// ---- SelfTests/TestCases/TestSuite_CommandAdapter/Test_CommandAdapterInitialization.TcPOU
{region 'Documentation'}
(*!
<summary>Verifies command-only initialization before cyclic use and after a retained sample.</summary>
<description>
PrimeHistory selects the reinitialization case: one public adapter call establishes TRUE history
before Initialize. The other instance calls Initialize before its first-ever cyclic use.
Both variants seed every command and distinctive Name/Status values. Initialize must clear
commands without touching the projection or invoking owner requests. Two fresh samples then
prove the old history was discarded and normal forwarding still works. No Event Buffer is
bound to this request-only double or to the production adapter; buffer work is outside its API.
Repeat runs reinitialize the same instance before the next script, rather than claiming fresh
instance memory. Assertions use the outer selftest publisher; the subject has no publisher.
</description>
*)
{endregion}
FUNCTION_BLOCK Test_CommandAdapterInitialization EXTENDS TestCaseBase
VAR_INPUT
    PrimeHistory : BOOL := FALSE; //! TRUE primes one TRUE command sample before reinitialization; FALSE exercises first-ever initialization.
END_VAR
VAR
    FSubject : RunControlCommandAdapter;
    FOwner : RunControlRequestRecorder;
    FControl : ST_RunControl;
    FExpectedStatus : ST_RunControlStatus;
    FStep : UINT;
    FChecked : BOOL;
    FCommandsCleared : AssertTrue;
    FCommandsClearedMatches : BOOL;
    FProjectionPreserved : AssertTrue;
    FProjectionPreservedMatches : BOOL;
    FNoRequests : AssertTrue;
    FNoRequestsMatches : BOOL;
    FHistoryCleared : AssertTrue;
    FHistoryClearedMatches : BOOL;
    FFreshRequest : AssertTrue;
    FFreshRequestMatches : BOOL;
END_VAR
VAR CONSTANT
    InitializeSubject : UINT := 0;
    FirstSample : UINT := 1;
    SecondSample : UINT := 2;
    CheckResults : UINT := 3;
END_VAR

SUPER^();

{region 'Documentation'}
(*!
<summary>Collects the five independent initialization checks.</summary>
*)
{endregion}
METHOD PROTECTED AggregateResults
VAR_INPUT
    Aggregator : I_ResultAggregator; //! Borrowed result sink owned by the outer Test Case; add this test's checking Assertions without resetting or retaining the sink.
END_VAR
Aggregator.AddProvider(Provider := FCommandsCleared);
Aggregator.AddProvider(Provider := FProjectionPreserved);
Aggregator.AddProvider(Provider := FNoRequests);
Aggregator.AddProvider(Provider := FHistoryCleared);
Aggregator.AddProvider(Provider := FFreshRequest);
END_METHOD

{region 'Documentation'}
(*!
<summary>Configures one scripted initialization test and its checking Assertions.</summary>
*)
{endregion}
METHOD PROTECTED Configure
FPreparationStateCount := 0;
FTestStateCount := 1;
FCommandsCleared.Initialize(Parent := THIS^,
    AssertionName := 'CommandsCleared');
FProjectionPreserved.Initialize(Parent := THIS^,
    AssertionName := 'ProjectionPreserved');
FNoRequests.Initialize(Parent := THIS^,
    AssertionName := 'NoRequests');
FHistoryCleared.Initialize(Parent := THIS^,
    AssertionName := 'HistoryCleared');
FFreshRequest.Initialize(Parent := THIS^,
    AssertionName := 'FreshRequest');
END_METHOD

{region 'Documentation'}
(*!
<summary>No asynchronous resource needs abort processing.</summary>
*)
{endregion}
METHOD PROTECTED ProcessAbort
VAR_INPUT
    Enable : BOOL; //! Phase permission supplied by the owning Test Case; FALSE does not authorize progression, while observation may continue.
END_VAR
IF Enable THEN
    CompleteAbort();
END_IF;
END_METHOD

{region 'Documentation'}
(*!
<summary>Evaluates stored observations after the bounded three-step script.</summary>
*)
{endregion}
METHOD PROTECTED ProcessAssertions
VAR_INPUT
    Enable : BOOL; //! Phase permission supplied by the owning Test Case; FALSE does not authorize progression, while observation may continue.
END_VAR
VAR
    Evaluate : BOOL;
END_VAR
Evaluate := Enable AND (FStep = CheckResults);
FCommandsCleared(Enable := Evaluate,
    State := State,
    IN := FCommandsClearedMatches);
FProjectionPreserved(Enable := Evaluate,
    State := State,
    IN := FProjectionPreservedMatches);
FNoRequests(Enable := Evaluate,
    State := State,
    IN := FNoRequestsMatches);
FHistoryCleared(Enable := Evaluate,
    State := State,
    IN := FHistoryClearedMatches);
FFreshRequest(Enable := Evaluate,
    State := State,
    IN := FFreshRequestMatches);
IF Evaluate THEN
    FChecked := TRUE;
END_IF;
END_METHOD

{region 'Documentation'}
(*!
<summary>No Preparation phase is needed.</summary>
*)
{endregion}
METHOD PROTECTED ProcessPreparations
VAR_INPUT
    // SA0033: Required override; this test has no Preparation work.
    {attribute 'analysis' := '-33'}
    Enable : BOOL; //! Phase permission supplied by the owning Test Case; FALSE does not authorize progression, while observation may continue.
END_VAR
END_METHOD

{region 'Documentation'}
(*!
<summary>Resets the test script; subject initialization remains the operation under test.</summary>
*)
{endregion}
METHOD PROTECTED ProcessReset
FStep := InitializeSubject;
FChecked := FALSE;
FOwner.Clear();
FCommandsCleared.Reset();
FCommandsClearedMatches := FALSE;
FProjectionPreserved.Reset();
FProjectionPreservedMatches := FALSE;
FNoRequests.Reset();
FNoRequestsMatches := FALSE;
FHistoryCleared.Reset();
FHistoryClearedMatches := FALSE;
FFreshRequest.Reset();
FFreshRequestMatches := FALSE;
CompleteReset();
END_METHOD

{region 'Documentation'}
(*!
<summary>Initializes before cyclic use, then checks history through two fresh samples.</summary>
*)
{endregion}
METHOD PROTECTED ProcessTests
VAR_INPUT
    Enable : BOOL; //! Phase permission supplied by the owning Test Case; FALSE does not authorize progression, while observation may continue.
END_VAR
IF NOT Enable THEN
    RETURN;
END_IF;
IF FChecked THEN
    CompleteTests();
    RETURN;
END_IF;
CASE FStep OF
    InitializeSubject:
        SeedControl();
        FOwner.Clear();
        IF PrimeHistory THEN
            // Establish stale TRUE samples through the public call, never by editing private history.
            FSubject(RunControl := FOwner,
                Commands := FControl.Cmd);
            FNoRequestsMatches := (FOwner.StartCount = 0) AND (FOwner.AbortCount = 0) AND (FOwner.ResetCount = 0);
        ELSE
            FNoRequestsMatches := TRUE;
        END_IF;
        FSubject.Initialize(ControlData := FControl);
        FCommandsClearedMatches := NOT FControl.Cmd.Start AND NOT FControl.Cmd.Abort AND NOT FControl.Cmd.Reset
            AND NOT FControl.BufferCmd.Reset AND (FControl.BufferCmd.DeleteSequenceId = 0);
        FProjectionPreservedMatches := (FControl.Name = 'PreservedRoot')
            AND (FControl.Status.Execution.State = FExpectedStatus.Execution.State)
            AND (FControl.Status.Execution.ExecutionStatus = FExpectedStatus.Execution.ExecutionStatus)
            AND (FControl.Status.Execution.Result = FExpectedStatus.Execution.Result)
            AND (FControl.Status.Execution.Uninitialized = FExpectedStatus.Execution.Uninitialized)
            AND (FControl.Status.Execution.ConfigError = FExpectedStatus.Execution.ConfigError)
            AND (FControl.Status.Execution.Ready = FExpectedStatus.Execution.Ready)
            AND (FControl.Status.Execution.Running = FExpectedStatus.Execution.Running)
            AND (FControl.Status.Execution.Completed = FExpectedStatus.Execution.Completed)
            AND (FControl.Status.Execution.Aborted = FExpectedStatus.Execution.Aborted)
            AND (FControl.Status.Execution.Inactive = FExpectedStatus.Execution.Inactive)
            AND (FControl.Status.Execution.Error = FExpectedStatus.Execution.Error)
            AND (FControl.Status.SuiteCountTotal = FExpectedStatus.SuiteCountTotal)
            AND (FControl.Status.SuiteCountInactive = FExpectedStatus.SuiteCountInactive)
            AND (FControl.Status.SuiteCountIdle = FExpectedStatus.SuiteCountIdle)
            AND (FControl.Status.SuiteCountRunning = FExpectedStatus.SuiteCountRunning)
            AND (FControl.Status.SuiteCountCompleted = FExpectedStatus.SuiteCountCompleted)
            AND (FControl.Status.SuiteCountPassed = FExpectedStatus.SuiteCountPassed)
            AND (FControl.Status.SuiteCountFailed = FExpectedStatus.SuiteCountFailed)
            AND (FControl.Status.SuiteCountError = FExpectedStatus.SuiteCountError)
            AND (FControl.Status.Runtime = FExpectedStatus.Runtime);
        FNoRequestsMatches := FNoRequestsMatches AND (FOwner.StartCount = 0) AND (FOwner.AbortCount = 0) AND (FOwner.ResetCount = 0);
        FStep := FirstSample;
    FirstSample:
        FControl.Cmd.Start := TRUE;
        FControl.Cmd.Abort := TRUE;
        FControl.Cmd.Reset := TRUE;
        FSubject(RunControl := FOwner,
            Commands := FControl.Cmd);
        FHistoryClearedMatches := (FOwner.StartCount = 0) AND (FOwner.AbortCount = 0) AND (FOwner.ResetCount = 0)
            AND FControl.Cmd.Start AND FControl.Cmd.Abort AND FControl.Cmd.Reset;
        FStep := SecondSample;
    SecondSample:
        FSubject(RunControl := FOwner,
            Commands := FControl.Cmd);
        FFreshRequestMatches := (FOwner.StartCount = 1) AND (FOwner.AbortCount = 1)
            AND (FOwner.ResetCount = 1) AND NOT FControl.Cmd.Start AND NOT FControl.Cmd.Abort AND NOT FControl.Cmd.Reset;
        FStep := CheckResults;
END_CASE;
END_METHOD

{region 'Documentation'}
(*!
<summary>Uses distinctive projection sentinels, deliberately not a valid lifecycle snapshot.</summary>
*)
{endregion}
METHOD PRIVATE SeedControl
FControl.Name := 'PreservedRoot';
FControl.Status.Execution.State := E_State.Completed;
FControl.Status.Execution.ExecutionStatus := E_ExecutionStatus.Completed;
FControl.Status.Execution.Result := E_Result.Failed;
FControl.Status.Execution.Uninitialized := TRUE;
FControl.Status.Execution.ConfigError := TRUE;
FControl.Status.Execution.Ready := TRUE;
FControl.Status.Execution.Running := TRUE;
FControl.Status.Execution.Completed := TRUE;
FControl.Status.Execution.Aborted := TRUE;
FControl.Status.Execution.Inactive := TRUE;
FControl.Status.Execution.Error := TRUE;
FControl.Status.SuiteCountTotal := 1;
FControl.Status.SuiteCountInactive := 2;
FControl.Status.SuiteCountIdle := 3;
FControl.Status.SuiteCountRunning := 4;
FControl.Status.SuiteCountCompleted := 5;
FControl.Status.SuiteCountPassed := 6;
FControl.Status.SuiteCountFailed := 7;
FControl.Status.SuiteCountError := 8;
FControl.Status.Runtime := T#123ms;
FExpectedStatus := FControl.Status;
FControl.Cmd.Start := TRUE;
FControl.Cmd.Abort := TRUE;
FControl.Cmd.Reset := TRUE;
FControl.BufferCmd.Reset := TRUE;
FControl.BufferCmd.DeleteSequenceId := 123;
END_METHOD

END_FUNCTION_BLOCK

// ---- Framework/RunControl/POU/RunControlCommandAdapter.TcPOU
{region 'Documentation'}
(*!
<summary>Qualifies external lifecycle commands and forwards requests before the Run Control FB call.</summary>
<description>
Initialize with the selected ControlData at PLC startup before the first cyclic call.
Requires a valid Run Control interface and its actual command storage, with stable cyclic wiring.

Call once before the matching concrete Run Control in the same task. A lifecycle bit must be TRUE in two consecutive adapter samples before it is forwarded and cleared. Multiple accepted bits are all forwarded; Run Control later applies Reset over Abort over Start. Initialize clears both lifecycle and Buffer commands at startup, while regular calls handle only lifecycle bits. There is no null-interface check or automatic storage-identity validation; the application owns valid, stable wiring.
</description>
*)
{endregion}
FUNCTION_BLOCK RunControlCommandAdapter
VAR_INPUT
    // SA0027: Parameter denotes the supplied owner interface, not the concrete RunControl FB.
    {attribute 'analysis' := '-27'}
    RunControl : I_RunControl; //! Nonzero request recipient matching Commands storage; an uninitialized owner discards forwarded requests.
END_VAR
VAR_IN_OUT
    Commands : ST_Command; //! Actual external lifecycle-command storage; commands are qualified, forwarded and cleared in place.
END_VAR
VAR
    FPreviousCommands : ST_Command;
END_VAR

IF Commands.Reset AND FPreviousCommands.Reset THEN
    RunControl.RequestReset();
    Commands.Reset := FALSE;
END_IF;

IF Commands.Abort AND FPreviousCommands.Abort THEN
    RunControl.RequestAbort();
    Commands.Abort := FALSE;
END_IF;

IF Commands.Start AND FPreviousCommands.Start THEN
    RunControl.RequestStart();
    Commands.Start := FALSE;
END_IF;

FPreviousCommands := Commands;

{region 'Documentation'}
(*!
<summary>Clears external commands and sampling history once at PLC startup, before Event Buffer/hierarchy initialization.</summary>
<description>
Preserves Name and Status; does not use cyclic inputs, invoke requests or execute buffer operations.
</description>
*)
{endregion}
METHOD PUBLIC Initialize
VAR_IN_OUT
    ControlData : ST_RunControl; //! External Run Control storage; Initialize clears Cmd and BufferCmd without changing Name or Status.
END_VAR
ControlData.Cmd.Start := FALSE;
ControlData.Cmd.Abort := FALSE;
ControlData.Cmd.Reset := FALSE;
ControlData.BufferCmd.Reset := FALSE;
ControlData.BufferCmd.DeleteSequenceId := 0;

FPreviousCommands.Start := FALSE;
FPreviousCommands.Abort := FALSE;
FPreviousCommands.Reset := FALSE;
END_METHOD

END_FUNCTION_BLOCK

// ---- SelfTests/TestCases/TestSuite_CommandAdapter/Helper/RunControlRequestRecorder.TcPOU
{region 'Documentation'}
(*!
<summary>Request-only I_RunControl double; counts calls without simulating lifecycle behavior.</summary>
*)
{endregion}
FUNCTION_BLOCK RunControlRequestRecorder IMPLEMENTS I_RunControl
VAR
    FStartCount : UINT;
    FAbortCount : UINT;
    FResetCount : UINT;
    FStatus : ST_RunControlStatus;
END_VAR

{region 'Documentation'}
(*!
<summary>Passive AbortCount observation for the command-adapter tests.</summary>
*)
{endregion}
{attribute 'monitoring' := 'call'}
PROPERTY PUBLIC AbortCount : UINT //! Passive AbortCount observation for the command-adapter tests.
GET // PUBLIC
AbortCount := FAbortCount;
END_GET
END_PROPERTY

{region 'Documentation'}
(*!
<summary>Clears recorded calls without performing lifecycle work.</summary>
*)
{endregion}
METHOD PUBLIC Clear
FStartCount := 0;
FAbortCount := 0;
FResetCount := 0;
END_METHOD

{region 'Documentation'}
(*!
<summary>Passive Name observation for the command-adapter tests.</summary>
*)
{endregion}
{attribute 'monitoring' := 'variable'}
PROPERTY PUBLIC Name : STRING(GVL_Constants.NameLength) //! Passive Name observation for the command-adapter tests.
GET // PUBLIC
Name := 'CommandTarget';
END_GET
END_PROPERTY

{region 'Documentation'}
(*!
<summary>Records a Abort request only; no lifecycle or buffer operations.</summary>
*)
{endregion}
METHOD PUBLIC RequestAbort
FAbortCount := FAbortCount + 1;
END_METHOD

{region 'Documentation'}
(*!
<summary>Records a Reset request only; no lifecycle or buffer operations.</summary>
*)
{endregion}
METHOD PUBLIC RequestReset
FResetCount := FResetCount + 1;
END_METHOD

{region 'Documentation'}
(*!
<summary>Records a Start request only; no lifecycle or buffer operations.</summary>
*)
{endregion}
METHOD PUBLIC RequestStart
FStartCount := FStartCount + 1;
END_METHOD

{region 'Documentation'}
(*!
<summary>Passive ResetCount observation for the command-adapter tests.</summary>
*)
{endregion}
{attribute 'monitoring' := 'call'}
PROPERTY PUBLIC ResetCount : UINT //! Passive ResetCount observation for the command-adapter tests.
GET // PUBLIC
ResetCount := FResetCount;
END_GET
END_PROPERTY

{region 'Documentation'}
(*!
<summary>Passive Result observation for the command-adapter tests.</summary>
*)
{endregion}
{attribute 'monitoring' := 'call'}
PROPERTY PUBLIC Result : E_Result //! Passive Result observation for the command-adapter tests.
GET // PUBLIC
Result := E_Result.NotEvaluated;
END_GET
END_PROPERTY

{region 'Documentation'}
(*!
<summary>Passive StartCount observation for the command-adapter tests.</summary>
*)
{endregion}
{attribute 'monitoring' := 'call'}
PROPERTY PUBLIC StartCount : UINT //! Passive StartCount observation for the command-adapter tests.
GET // PUBLIC
StartCount := FStartCount;
END_GET
END_PROPERTY

{region 'Documentation'}
(*!
<summary>Passive Status observation for the command-adapter tests.</summary>
*)
{endregion}
PROPERTY PUBLIC Status : ST_RunControlStatus //! Passive Status observation for the command-adapter tests.
GET // PUBLIC
Status := FStatus;
END_GET
END_PROPERTY

END_FUNCTION_BLOCK

// ---- SelfTests/TestCases/TestSuite_CommandAdapter/Test_CommandQualification.TcPOU
{region 'Documentation'}
(*!
<summary>Checks two-sample qualification and PLC-owned clearing for one external lifecycle command.</summary>
<description>
Use one instance per Start, Abort and Reset. Every enabled cycle samples the real adapter once.
The script first withdraws two separate one-sample pulses, then leaves TRUE untouched for two
calls. Acceptance must forward exactly one request and clear that field. A following call
without a write must not repeat it. A new TRUE then needs two new samples before request two.
Each sample checks the selected count/bit and both unrelated commands. This is deterministic
call-boundary evidence, not a simulation of asynchronous ADS writes or a command handshake.
ProcessReset initializes the local subject and clears the recorder for repeatable runs.
</description>
*)
{endregion}
FUNCTION_BLOCK Test_CommandQualification EXTENDS TestCaseBase
VAR_INPUT
    Command : E_AdapterCommand := E_AdapterCommand.Start; //! External command field exercised by this instance; held fixed by the containing Suite.
END_VAR
VAR
    FSubject : RunControlCommandAdapter;
    FOwner : RunControlRequestRecorder;
    FControl : ST_RunControl;
    FStep : UINT;
    FSampleChecked : BOOL;
    FRequestCount : AssertTrue;
    FRequestCountMatches : BOOL;
    FCommandValue : AssertTrue;
    FCommandValueMatches : BOOL;
    FOtherCommands : AssertTrue;
    FOtherCommandsMatches : BOOL;
END_VAR
VAR CONSTANT
    Baseline : UINT := 0;
    SinglePulse : UINT := 1;
    Withdrawal : UINT := 2;
    SeparatedPulse : UINT := 3;
    SecondWithdrawal : UINT := 4;
    RetainedFirstSample : UINT := 5;
    RetainedSecondSample : UINT := 6;
    FreshFirstSample : UINT := 8;
    FreshSecondSample : UINT := 9;
    AfterFreshClearing : UINT := 10;
END_VAR

SUPER^();

{region 'Documentation'}
(*!
<summary>Collects request-count, field-value and isolation checks.</summary>
*)
{endregion}
METHOD PROTECTED AggregateResults
VAR_INPUT
    Aggregator : I_ResultAggregator; //! Borrowed result sink owned by the outer Test Case; add this test's checking Assertions without resetting or retaining the sink.
END_VAR
Aggregator.AddProvider(Provider := FRequestCount);
Aggregator.AddProvider(Provider := FCommandValue);
Aggregator.AddProvider(Provider := FOtherCommands);
END_METHOD

{region 'Documentation'}
(*!
<summary>Checks the explicit script oracle against recorded calls and the post-call command fields.</summary>
*)
{endregion}
METHOD PRIVATE CheckSample
VAR
    ExpectedCount : UINT;
    ExpectedCommand : BOOL;
    ActualCount : UINT;
    ActualCommand : BOOL;
END_VAR
IF FStep >= FreshSecondSample THEN
    ExpectedCount := 2;
ELSIF FStep >= RetainedSecondSample THEN
    ExpectedCount := 1;
END_IF;
ExpectedCommand := (FStep = SinglePulse) OR (FStep = SeparatedPulse)
    OR (FStep = RetainedFirstSample) OR (FStep = FreshFirstSample);
CASE Command OF
    E_AdapterCommand.Start:
        ActualCount := FOwner.StartCount;
        ActualCommand := FControl.Cmd.Start;
        FOtherCommandsMatches := (FOwner.AbortCount = 0) AND (FOwner.ResetCount = 0)
            AND NOT FControl.Cmd.Abort AND NOT FControl.Cmd.Reset;
    E_AdapterCommand.Abort:
        ActualCount := FOwner.AbortCount;
        ActualCommand := FControl.Cmd.Abort;
        FOtherCommandsMatches := (FOwner.StartCount = 0) AND (FOwner.ResetCount = 0)
            AND NOT FControl.Cmd.Start AND NOT FControl.Cmd.Reset;
    E_AdapterCommand.Reset:
        ActualCount := FOwner.ResetCount;
        ActualCommand := FControl.Cmd.Reset;
        FOtherCommandsMatches := (FOwner.StartCount = 0) AND (FOwner.AbortCount = 0)
            AND NOT FControl.Cmd.Start AND NOT FControl.Cmd.Abort;
END_CASE;
FRequestCountMatches := ActualCount = ExpectedCount;
FCommandValueMatches := ActualCommand = ExpectedCommand;
END_METHOD

{region 'Documentation'}
(*!
<summary>Initializes the three checking Assertions for the selected command.</summary>
*)
{endregion}
METHOD PROTECTED Configure
FPreparationStateCount := 0;
FTestStateCount := 1;
FRequestCount.Initialize(Parent := THIS^,
    AssertionName := 'RequestCount');
FCommandValue.Initialize(Parent := THIS^,
    AssertionName := 'CommandValue');
FOtherCommands.Initialize(Parent := THIS^,
    AssertionName := 'OtherCommands');
END_METHOD

{region 'Documentation'}
(*!
<summary>No asynchronous resource needs abort handling.</summary>
*)
{endregion}
METHOD PROTECTED ProcessAbort
VAR_INPUT
    Enable : BOOL; //! Phase permission supplied by the owning Test Case; FALSE does not authorize progression, while observation may continue.
END_VAR
IF Enable THEN
    CompleteAbort();
END_IF;
END_METHOD

{region 'Documentation'}
(*!
<summary>Checks every sample before advancing; failures remain latched across the script.</summary>
*)
{endregion}
METHOD PROTECTED ProcessAssertions
VAR_INPUT
    Enable : BOOL; //! Phase permission supplied by the owning Test Case; FALSE does not authorize progression, while observation may continue.
END_VAR
FRequestCount(Enable := Enable,
    State := State,
    IN := FRequestCountMatches);
FCommandValue(Enable := Enable,
    State := State,
    IN := FCommandValueMatches);
FOtherCommands(Enable := Enable,
    State := State,
    IN := FOtherCommandsMatches);
IF Enable THEN
    FSampleChecked := TRUE;
END_IF;
END_METHOD

{region 'Documentation'}
(*!
<summary>No Preparation work is required.</summary>
*)
{endregion}
METHOD PROTECTED ProcessPreparations
VAR_INPUT
    // SA0033: Required override; this test has no Preparation phase.
    {attribute 'analysis' := '-33'}
    Enable : BOOL; //! Phase permission supplied by the owning Test Case; FALSE does not authorize progression, while observation may continue.
END_VAR
END_METHOD

{region 'Documentation'}
(*!
<summary>Clears subject history, recorded requests and the bounded sample script.</summary>
*)
{endregion}
METHOD PROTECTED ProcessReset
FSubject.Initialize(ControlData := FControl);
FOwner.Clear();
FStep := Baseline;
FSampleChecked := FALSE;
FRequestCount.Reset();
FRequestCountMatches := FALSE;
FCommandValue.Reset();
FCommandValueMatches := FALSE;
FOtherCommands.Reset();
FOtherCommandsMatches := FALSE;
CompleteReset();
END_METHOD

{region 'Documentation'}
(*!
<summary>Applies one scheduled write and one real adapter call per active PLC cycle.</summary>
*)
{endregion}
METHOD PROTECTED ProcessTests
VAR_INPUT
    Enable : BOOL; //! Phase permission supplied by the owning Test Case; FALSE does not authorize progression, while observation may continue.
END_VAR
IF NOT Enable THEN
    RETURN;
END_IF;
IF FSampleChecked THEN
    IF FStep = AfterFreshClearing THEN
        CompleteTests();
        RETURN;
    END_IF;
    FStep := FStep + 1;
    FSampleChecked := FALSE;
END_IF;
CASE FStep OF
    SinglePulse, SeparatedPulse, RetainedFirstSample, FreshFirstSample:
        SetCommand(Value := TRUE);
    Withdrawal, SecondWithdrawal:
        SetCommand(Value := FALSE);
ELSE
    // No external write: retain the actual field, including the adapter's clearing.
END_CASE;
FSubject(RunControl := FOwner,
    Commands := FControl.Cmd);
CheckSample();
END_METHOD

{region 'Documentation'}
(*!
<summary>Writes only the chosen external command field.</summary>
*)
{endregion}
METHOD PRIVATE SetCommand
VAR_INPUT
    Value : BOOL; //! Boolean value written only to the selected command field.
END_VAR
CASE Command OF
    E_AdapterCommand.Start:
        FControl.Cmd.Start := Value;
    E_AdapterCommand.Abort:
        FControl.Cmd.Abort := Value;
    E_AdapterCommand.Reset:
        FControl.Cmd.Reset := Value;
END_CASE;
END_METHOD

END_FUNCTION_BLOCK

// ---- SelfTests/TestCases/TestSuite_CommandAdapter/Test_CommandIndependence.TcPOU
{region 'Documentation'}
(*!
<summary>Verifies independent command qualification and selective clearing across staggered writes.</summary>
<description>
The initial Start/Reset pair is sampled before Abort is written after that call. The pair
must be forwarded while Abort remains pending. Further post-call Start, Reset and Abort
writes rotate which field is newly sampled versus accepted. After those requests drain,
all three bits are raised together and must all be forwarded exactly once after two samples.
Fixed count and bit traces are the oracle; no request order or lifecycle priority is asserted.
Buffer commands and selected Name/Status fields are changed before each call and must survive.
CheckSample captures pre-post-write observations so Assertion processing cannot confuse the
test's own later writes with the adapter's output. There is one subject call per active cycle.
These deterministic boundaries do not prove arbitrary ADS interleavings inside an FB call.
</description>
*)
{endregion}
FUNCTION_BLOCK Test_CommandIndependence EXTENDS TestCaseBase
VAR
    FSubject : RunControlCommandAdapter;
    FOwner : RunControlRequestRecorder;
    FControl : ST_RunControl;
    FStep : UINT;
    FSampleChecked : BOOL;
    FForwarding : AssertTrue;
    FForwardingMatches : BOOL;
    FSelectiveClearing : AssertTrue;
    FSelectiveClearingMatches : BOOL;
    FUnrelatedFields : AssertTrue;
    FUnrelatedFieldsMatches : BOOL;
END_VAR
VAR CONSTANT
    PairFirstSample : UINT := 0;
    PairAccepted : UINT := 1;
    AbortAccepted : UINT := 2;
    StartAccepted : UINT := 3;
    ResetAccepted : UINT := 4;
    SecondAbortAccepted : UINT := 5;
    AllFirstSample : UINT := 8;
    LastSample : UINT := 10;
    ExpectedStartCounts : ARRAY[0..LastSample] OF UINT := [0, 1, 1, 2, 2, 2, 3, 3, 3, 4, 4];
    ExpectedAbortCounts : ARRAY[0..LastSample] OF UINT := [0, 0, 1, 1, 1, 2, 2, 2, 2, 3, 3];
    ExpectedResetCounts : ARRAY[0..LastSample] OF UINT := [0, 1, 1, 1, 2, 2, 2, 3, 3, 4, 4];
    ExpectedStartBits : ARRAY[0..LastSample] OF BOOL := [TRUE, FALSE, TRUE, FALSE, FALSE, TRUE, FALSE, FALSE, TRUE, FALSE, FALSE];
    ExpectedAbortBits : ARRAY[0..LastSample] OF BOOL := [FALSE, TRUE, FALSE, FALSE, TRUE, FALSE, FALSE, FALSE, TRUE, FALSE, FALSE];
    ExpectedResetBits : ARRAY[0..LastSample] OF BOOL := [TRUE, FALSE, FALSE, TRUE, FALSE, FALSE, TRUE, FALSE, TRUE, FALSE, FALSE];
END_VAR

SUPER^();

{region 'Documentation'}
(*!
<summary>Collects only the checking Assertions.</summary>
*)
{endregion}
METHOD PROTECTED AggregateResults
VAR_INPUT
    Aggregator : I_ResultAggregator; //! Borrowed result sink owned by the outer Test Case; add this test's checking Assertions without resetting or retaining the sink.
END_VAR
Aggregator.AddProvider(Provider := FForwarding);
Aggregator.AddProvider(Provider := FSelectiveClearing);
Aggregator.AddProvider(Provider := FUnrelatedFields);
END_METHOD

{region 'Documentation'}
(*!
<summary>Uses fixed expected traces, independent of adapter request order.</summary>
*)
{endregion}
METHOD PRIVATE CheckSample
FForwardingMatches := (FOwner.StartCount = ExpectedStartCounts[FStep])
    AND (FOwner.AbortCount = ExpectedAbortCounts[FStep])
    AND (FOwner.ResetCount = ExpectedResetCounts[FStep]);
FSelectiveClearingMatches := (FControl.Cmd.Start = ExpectedStartBits[FStep])
    AND (FControl.Cmd.Abort = ExpectedAbortBits[FStep])
    AND (FControl.Cmd.Reset = ExpectedResetBits[FStep]);
FUnrelatedFieldsMatches := (FControl.Name = 'CommandProjection')
    AND (FControl.Status.Execution.State = E_State.Completed)
    AND (FControl.Status.Execution.Result = E_Result.Failed)
    AND (FControl.Status.SuiteCountTotal = FStep + 1)
    AND (FControl.Status.Runtime = UINT_TO_TIME(FStep + 1))
    AND (FControl.BufferCmd.Reset = ((FStep MOD 2) = 0))
    AND (FControl.BufferCmd.DeleteSequenceId = UINT_TO_UDINT(FStep + 1));
END_METHOD

{region 'Documentation'}
(*!
<summary>Initializes the independent forwarding, clearing and projection checks.</summary>
*)
{endregion}
METHOD PROTECTED Configure
FPreparationStateCount := 0;
FTestStateCount := 1;
FForwarding.Initialize(Parent := THIS^,
    AssertionName := 'Forwarding');
FSelectiveClearing.Initialize(Parent := THIS^,
    AssertionName := 'SelectiveClearing');
FUnrelatedFields.Initialize(Parent := THIS^,
    AssertionName := 'UnrelatedFields');
END_METHOD

{region 'Documentation'}
(*!
<summary>No asynchronous resource is involved.</summary>
*)
{endregion}
METHOD PROTECTED ProcessAbort
VAR_INPUT
    Enable : BOOL; //! Phase permission supplied by the owning Test Case; FALSE does not authorize progression, while observation may continue.
END_VAR
IF Enable THEN
    CompleteAbort();
END_IF;
END_METHOD

{region 'Documentation'}
(*!
<summary>Latches every sample's observations before the script advances.</summary>
*)
{endregion}
METHOD PROTECTED ProcessAssertions
VAR_INPUT
    Enable : BOOL; //! Phase permission supplied by the owning Test Case; FALSE does not authorize progression, while observation may continue.
END_VAR
FForwarding(Enable := Enable,
    State := State,
    IN := FForwardingMatches);
FSelectiveClearing(Enable := Enable,
    State := State,
    IN := FSelectiveClearingMatches);
FUnrelatedFields(Enable := Enable,
    State := State,
    IN := FUnrelatedFieldsMatches);
IF Enable THEN
    FSampleChecked := TRUE;
END_IF;
END_METHOD

{region 'Documentation'}
(*!
<summary>No Preparation phase is required.</summary>
*)
{endregion}
METHOD PROTECTED ProcessPreparations
VAR_INPUT
    // SA0033: Required override; this test has no Preparation phase.
    {attribute 'analysis' := '-33'}
    Enable : BOOL; //! Phase permission supplied by the owning Test Case; FALSE does not authorize progression, while observation may continue.
END_VAR
END_METHOD

{region 'Documentation'}
(*!
<summary>Clears local commands, sampling history, recorded calls and checking state.</summary>
*)
{endregion}
METHOD PROTECTED ProcessReset
FSubject.Initialize(ControlData := FControl);
FOwner.Clear();
FStep := PairFirstSample;
FSampleChecked := FALSE;
FForwarding.Reset();
FForwardingMatches := FALSE;
FSelectiveClearing.Reset();
FSelectiveClearingMatches := FALSE;
FUnrelatedFields.Reset();
FUnrelatedFieldsMatches := FALSE;
CompleteReset();
END_METHOD

{region 'Documentation'}
(*!
<summary>Places writes before or after one adapter call; captures observations before post-call writes.</summary>
*)
{endregion}
METHOD PROTECTED ProcessTests
VAR_INPUT
    Enable : BOOL; //! Phase permission supplied by the owning Test Case; FALSE does not authorize progression, while observation may continue.
END_VAR
IF NOT Enable THEN
    RETURN;
END_IF;
IF FSampleChecked THEN
    IF FStep = LastSample THEN
        CompleteTests();
        RETURN;
    END_IF;
    FStep := FStep + 1;
    FSampleChecked := FALSE;
END_IF;
CASE FStep OF
    PairFirstSample:
        FControl.Cmd.Start := TRUE;
        FControl.Cmd.Reset := TRUE;
    AllFirstSample:
        FControl.Cmd.Start := TRUE;
        FControl.Cmd.Abort := TRUE;
        FControl.Cmd.Reset := TRUE;
END_CASE;
FControl.Name := 'CommandProjection';
FControl.Status.Execution.State := E_State.Completed;
FControl.Status.Execution.Result := E_Result.Failed;
FControl.Status.SuiteCountTotal := FStep + 1;
FControl.Status.Runtime := UINT_TO_TIME(FStep + 1);
FControl.BufferCmd.Reset := (FStep MOD 2) = 0;
FControl.BufferCmd.DeleteSequenceId := UINT_TO_UDINT(FStep + 1);
FSubject(RunControl := FOwner,
    Commands := FControl.Cmd);
CheckSample();
// These writes happen after the observation and become the next call's first sample.
CASE FStep OF
    PairFirstSample, StartAccepted:
        FControl.Cmd.Abort := TRUE;
    PairAccepted, ResetAccepted:
        FControl.Cmd.Start := TRUE;
    AbortAccepted, SecondAbortAccepted:
        FControl.Cmd.Reset := TRUE;
END_CASE;
END_METHOD

END_FUNCTION_BLOCK

// ---- SelfTests/TestSuites/TestSuite_EventDelivery.TcPOU
{region 'Documentation'}
(*!
<summary>Groups isolated event storage, delivery and deletion-watermark tests.</summary>
*)
{endregion}
FUNCTION_BLOCK TestSuite_EventDelivery EXTENDS TestSuiteBase
VAR
    FStorageBinding : Test_EventStorageBinding;
    FContent : Test_EventContent;
    FBufferFull : Test_EventBufferFull;
    FRingOrder : Test_EventRingOrder;
    FDeleteWatermarks : Test_EventDeleteWatermarks;
    FDeleteWrappedFull : Test_EventDeleteWrappedFull;
    FDeleteLostSequence : Test_EventDeleteLostSequence;
    FDeleteCommandBoundary : Test_EventDeleteCommandBoundary;
    FTestCases : ARRAY[1..TestCaseCapacity] OF I_TestCase;
END_VAR
VAR CONSTANT
    TestCaseCapacity : UINT := 8;
END_VAR

SUPER^();

{region 'Documentation'}
(*!
<summary>Initializes and registers the isolated event scenarios for serial execution.</summary>
*)
{endregion}
METHOD PROTECTED Configure
VAR_IN_OUT
    // SA0167: Borrowed owner builder; no temporary instance is created.
    {attribute 'analysis' := '-167'}
    Builder : TestSuiteConfigurationBuilder; //! Borrowed owner configuration builder used only during this Configure call; register this owner's concrete children.
END_VAR
VAR
    TestConfig : ST_TestCaseConfig;
END_VAR
Builder.Initialize(Mode := E_OrchestrationMode.Serial,
    TestCases := FTestCases);
FStorageBinding.Initialize(Parent := THIS^,
    TestName := 'StorageBinding',
    Config := TestConfig);
Builder.Register(TestCase := FStorageBinding);
FContent.Initialize(Parent := THIS^,
    TestName := 'Content',
    Config := TestConfig);
Builder.Register(TestCase := FContent);
FBufferFull.Initialize(Parent := THIS^,
    TestName := 'BufferFull',
    Config := TestConfig);
Builder.Register(TestCase := FBufferFull);
FRingOrder.Initialize(Parent := THIS^,
    TestName := 'RingOrder',
    Config := TestConfig);
Builder.Register(TestCase := FRingOrder);
FDeleteWatermarks.Initialize(Parent := THIS^,
    TestName := 'DeleteWatermarks',
    Config := TestConfig);
Builder.Register(TestCase := FDeleteWatermarks);
FDeleteWrappedFull.Initialize(Parent := THIS^,
    TestName := 'DeleteWrappedFull',
    Config := TestConfig);
Builder.Register(TestCase := FDeleteWrappedFull);
FDeleteLostSequence.Initialize(Parent := THIS^,
    TestName := 'DeleteLostSequence',
    Config := TestConfig);
Builder.Register(TestCase := FDeleteLostSequence);
FDeleteCommandBoundary.Initialize(Parent := THIS^,
    TestName := 'DeleteCommandBoundary',
    Config := TestConfig);
Builder.Register(TestCase := FDeleteCommandBoundary);
END_METHOD

{region 'Documentation'}
(*!
<summary>Returns a registered scenario using its original array index.</summary>
*)
{endregion}
METHOD PUBLIC GetTestCase : I_TestCase //! Typed child interface at the original array index; zero when no entry is available.
VAR_INPUT
    Index : DINT; //! Original occupied child-array index, rather than an ordinal position.
END_VAR
GetTestCase := 0;
IF (ChildCount = 0) OR (Index < ChildArrayLowerBound)
    OR (DINT_TO_LINT(Index) >= DINT_TO_LINT(ChildArrayLowerBound) + UINT_TO_LINT(ChildCount)) THEN
    RETURN;
END_IF;
GetTestCase := FTestCases[Index];
END_METHOD

{region 'Documentation'}
(*!
<summary>Calls each owned scenario once per initialized Suite cycle.</summary>
*)
{endregion}
METHOD PROTECTED ProcessTestCases
FStorageBinding();
FContent();
FBufferFull();
FRingOrder();
FDeleteWatermarks();
FDeleteWrappedFull();
FDeleteLostSequence();
FDeleteCommandBoundary();
END_METHOD

END_FUNCTION_BLOCK

// ---- SelfTests/TestCases/TestSuite_EventDelivery/Test_EventStorageBinding.TcPOU
{region 'Documentation'}
(*!
<summary>Verifies two real Event Buffers publish into their own bound arrays and status structures.</summary>
<description>
The subjects own no global stream: each binds a static local array and separate projections.
Eight and twelve physical entries provide seven and eleven usable FIFO slots. One distinctive
event is published to each subject; observations are captured before the next operation so
cross-writes cannot be hidden by later initialization. The outer test Assertions use the
normal selftest publisher, which is never replaced. Every test run initializes both subjects
again; no production algorithm is copied and no private field is modified.
</description>
*)
{endregion}
FUNCTION_BLOCK Test_EventStorageBinding EXTENDS TestCaseBase
VAR
    FSmallBuffer : EventBuffer;
    FLargeBuffer : EventBuffer;
    FSmallEvents : ARRAY[1..SmallBufferLength] OF ST_Event;
    FLargeEvents : ARRAY[1..LargeBufferLength] OF ST_Event;
    FSmallFifo : ST_FifoStatus;
    FLargeFifo : ST_FifoStatus;
    FSmallStatus : ST_EventBufferStatus;
    FLargeStatus : ST_EventBufferStatus;
    FPerformed : BOOL;
    FChecked : BOOL;
    FBinding : AssertTrue;
    FBindingMatches : BOOL;
    FCapacity : AssertTrue;
    FCapacityMatches : BOOL;
    FInitialProjection : AssertTrue;
    FInitialProjectionMatches : BOOL;
    FSmallPublication : AssertTrue;
    FSmallPublicationMatches : BOOL;
    FLargePublication : AssertTrue;
    FLargePublicationMatches : BOOL;
    FIsolation : AssertTrue;
    FIsolationMatches : BOOL;
END_VAR
VAR CONSTANT
    SmallBufferLength : UINT := 8;
    LargeBufferLength : UINT := 12;
END_VAR

SUPER^();

{region 'Documentation'}
(*!
<summary>Collects the six independent storage-binding observations.</summary>
*)
{endregion}
METHOD PROTECTED AggregateResults
VAR_INPUT
    Aggregator : I_ResultAggregator; //! Borrowed result sink owned by the outer Test Case; add this test's checking Assertions without resetting or retaining the sink.
END_VAR
Aggregator.AddProvider(Provider := FBinding);
Aggregator.AddProvider(Provider := FCapacity);
Aggregator.AddProvider(Provider := FInitialProjection);
Aggregator.AddProvider(Provider := FSmallPublication);
Aggregator.AddProvider(Provider := FLargePublication);
Aggregator.AddProvider(Provider := FIsolation);
END_METHOD

{region 'Documentation'}
(*!
<summary>Requires successful initialization of all checking Assertions.</summary>
*)
{endregion}
METHOD PROTECTED CheckInitialization : BOOL //! TRUE when the inherited initialization check and this concrete fixture check both accept the setup.
CheckInitialization := FALSE;
IF NOT SUPER^.CheckInitialization() THEN
    RETURN;
END_IF;

CheckInitialization := FBinding.IsInitialized
    AND FCapacity.IsInitialized
    AND FInitialProjection.IsInitialized
    AND FSmallPublication.IsInitialized
    AND FLargePublication.IsInitialized
    AND FIsolation.IsInitialized;
END_METHOD

{region 'Documentation'}
(*!
<summary>Configures the single storage-binding scenario and its six Assertions.</summary>
*)
{endregion}
METHOD PROTECTED Configure
FPreparationStateCount := 0;
FTestStateCount := 1;
FBinding.Initialize(Parent := THIS^,
    AssertionName := 'Binding');
FCapacity.Initialize(Parent := THIS^,
    AssertionName := 'Capacity');
FInitialProjection.Initialize(Parent := THIS^,
    AssertionName := 'InitialProjection');
FSmallPublication.Initialize(Parent := THIS^,
    AssertionName := 'SmallPublication');
FLargePublication.Initialize(Parent := THIS^,
    AssertionName := 'LargePublication');
FIsolation.Initialize(Parent := THIS^,
    AssertionName := 'Isolation');
END_METHOD

{region 'Documentation'}
(*!
<summary>Binds differently sized static arrays and verifies initial projection and usable capacity.</summary>
*)
{endregion}
METHOD PRIVATE InitializeBuffers
VAR
    SmallInitialized : BOOL;
    LargeInitialized : BOOL;
    Index : UINT;
END_VAR
SmallInitialized := FSmallBuffer.Initialize(Buffer := FSmallEvents,
    FifoControl := FSmallFifo,
    Status := FSmallStatus);
LargeInitialized := FLargeBuffer.Initialize(Buffer := FLargeEvents,
    FifoControl := FLargeFifo,
    Status := FLargeStatus);
FBindingMatches := SmallInitialized AND LargeInitialized
    AND FSmallBuffer.IsValid AND FLargeBuffer.IsValid;
FCapacityMatches := (FSmallBuffer.Capacity = SmallBufferLength - 1)
    AND (FLargeBuffer.Capacity = LargeBufferLength - 1)
    AND (FSmallFifo.BufferLength = SmallBufferLength)
    AND (FLargeFifo.BufferLength = LargeBufferLength);
FInitialProjectionMatches := FSmallFifo.BufferEmpty AND FLargeFifo.BufferEmpty
    AND NOT FSmallFifo.ConfigError AND NOT FLargeFifo.ConfigError
    AND NOT FSmallFifo.IndexError AND NOT FLargeFifo.IndexError
    AND (FSmallFifo.ElementCount = 0) AND (FLargeFifo.ElementCount = 0)
    AND (FSmallFifo.IndexIn = 1) AND (FSmallFifo.IndexOut = 1)
    AND (FLargeFifo.IndexIn = 1) AND (FLargeFifo.IndexOut = 1)
    AND (FSmallStatus.SequenceId = 0) AND (FLargeStatus.SequenceId = 0)
    AND (FSmallStatus.DeletedSequenceId = 0) AND (FLargeStatus.DeletedSequenceId = 0)
    AND (FSmallStatus.LostEventCount = 0) AND (FLargeStatus.LostEventCount = 0);
FOR Index := 1 TO SmallBufferLength DO
    FInitialProjectionMatches := FInitialProjectionMatches AND (FSmallEvents[Index].SequenceId = 0);
END_FOR;
FOR Index := 1 TO LargeBufferLength DO
    FInitialProjectionMatches := FInitialProjectionMatches AND (FLargeEvents[Index].SequenceId = 0);
END_FOR;
END_METHOD

{region 'Documentation'}
(*!
<summary>Completes abort without asynchronous resource work.</summary>
*)
{endregion}
METHOD PROTECTED ProcessAbort
VAR_INPUT
    Enable : BOOL; //! Phase permission supplied by the owning Test Case; FALSE does not authorize progression, while observation may continue.
END_VAR
IF Enable THEN
    CompleteAbort();
END_IF;
END_METHOD

{region 'Documentation'}
(*!
<summary>Evaluates observations only after the two subjects have been exercised.</summary>
*)
{endregion}
METHOD PROTECTED ProcessAssertions
VAR_INPUT
    Enable : BOOL; //! Phase permission supplied by the owning Test Case; FALSE does not authorize progression, while observation may continue.
END_VAR
VAR
    Evaluate : BOOL;
END_VAR
Evaluate := Enable AND FPerformed;
FBinding(Enable := Evaluate,
    State := State,
    IN := FBindingMatches);
FCapacity(Enable := Evaluate,
    State := State,
    IN := FCapacityMatches);
FInitialProjection(Enable := Evaluate,
    State := State,
    IN := FInitialProjectionMatches);
FSmallPublication(Enable := Evaluate,
    State := State,
    IN := FSmallPublicationMatches);
FLargePublication(Enable := Evaluate,
    State := State,
    IN := FLargePublicationMatches);
FIsolation(Enable := Evaluate,
    State := State,
    IN := FIsolationMatches);
IF Evaluate THEN
    FChecked := TRUE;
END_IF;
END_METHOD

{region 'Documentation'}
(*!
<summary>No Preparation phase is needed.</summary>
*)
{endregion}
METHOD PROTECTED ProcessPreparations
VAR_INPUT
    // SA0033: Required override; this test has no Preparation work.
    {attribute 'analysis' := '-33'}
    Enable : BOOL; //! Phase permission supplied by the owning Test Case; FALSE does not authorize progression, while observation may continue.
END_VAR
END_METHOD

{region 'Documentation'}
(*!
<summary>Clears observations and Assertions; subject initialization remains under test.</summary>
*)
{endregion}
METHOD PROTECTED ProcessReset
FPerformed := FALSE;
FChecked := FALSE;
FBinding.Reset();
FBindingMatches := FALSE;
FCapacity.Reset();
FCapacityMatches := FALSE;
FInitialProjection.Reset();
FInitialProjectionMatches := FALSE;
FSmallPublication.Reset();
FSmallPublicationMatches := FALSE;
FLargePublication.Reset();
FLargePublicationMatches := FALSE;
FIsolation.Reset();
FIsolationMatches := FALSE;
CompleteReset();
END_METHOD

{region 'Documentation'}
(*!
<summary>Initializes and exercises the local bindings once per test run.</summary>
*)
{endregion}
METHOD PROTECTED ProcessTests
VAR_INPUT
    Enable : BOOL; //! Phase permission supplied by the owning Test Case; FALSE does not authorize progression, while observation may continue.
END_VAR
IF NOT Enable THEN
    RETURN;
END_IF;
IF FChecked THEN
    CompleteTests();
    RETURN;
END_IF;

IF NOT FPerformed THEN
    InitializeBuffers();
    PublishToSmallBuffer();
    PublishToLargeBuffer();
    FPerformed := TRUE;
END_IF;
END_METHOD

{region 'Documentation'}
(*!
<summary>Checks the second publication leaves the first buffer and its projections unchanged.</summary>
*)
{endregion}
METHOD PRIVATE PublishToLargeBuffer
VAR
    WriteResult : INT;
    Index : UINT;
END_VAR
WriteResult := FLargeBuffer.PublishEvent(Event := CreateFrameworkEvent(Name := 'LocalLarge',
    State := E_State.Idle,
    Severity := E_EventSeverity.Info,
    Message := 'Large binding'));
FLargePublicationMatches := (WriteResult = 1)
    AND (FLargeEvents[1].SequenceId = 1)
    AND (FLargeEvents[1].Name = 'LocalLarge') AND (FLargeEvents[1].Message = 'Large binding')
    AND (FLargeFifo.IndexIn = 2) AND (FLargeFifo.IndexOut = 1)
    AND (FLargeFifo.ElementCount = 1) AND NOT FLargeFifo.BufferEmpty
    AND (FLargeStatus.SequenceId = 1) AND (FLargeStatus.DeletedSequenceId = 0)
    AND (FLargeStatus.LostEventCount = 0);
FIsolationMatches := FIsolationMatches
    AND (FSmallEvents[1].SequenceId = 1)
    AND (FSmallEvents[1].Name = 'LocalSmall') AND (FSmallEvents[1].Message = 'Small binding')
    AND (FSmallFifo.IndexIn = 2) AND (FSmallFifo.IndexOut = 1)
    AND (FSmallFifo.ElementCount = 1) AND NOT FSmallFifo.BufferEmpty
    AND (FSmallStatus.SequenceId = 1) AND (FSmallStatus.DeletedSequenceId = 0)
    AND (FSmallStatus.LostEventCount = 0);
FOR Index := 2 TO SmallBufferLength DO
    FIsolationMatches := FIsolationMatches AND (FSmallEvents[Index].SequenceId = 0);
END_FOR;
END_METHOD

{region 'Documentation'}
(*!
<summary>Checks immediate local publication and that the other buffer is still empty.</summary>
*)
{endregion}
METHOD PRIVATE PublishToSmallBuffer
VAR
    WriteResult : INT;
    Index : UINT;
END_VAR
WriteResult := FSmallBuffer.PublishEvent(Event := CreateFrameworkEvent(Name := 'LocalSmall',
    State := E_State.Idle,
    Severity := E_EventSeverity.Info,
    Message := 'Small binding'));
FSmallPublicationMatches := (WriteResult = 1)
    AND (FSmallEvents[1].SequenceId = 1)
    AND (FSmallEvents[1].Name = 'LocalSmall') AND (FSmallEvents[1].Message = 'Small binding')
    AND (FSmallFifo.IndexIn = 2) AND (FSmallFifo.IndexOut = 1)
    AND (FSmallFifo.ElementCount = 1) AND NOT FSmallFifo.BufferEmpty
    AND (FSmallStatus.SequenceId = 1) AND (FSmallStatus.DeletedSequenceId = 0)
    AND (FSmallStatus.LostEventCount = 0);
FIsolationMatches := FLargeFifo.BufferEmpty AND (FLargeFifo.ElementCount = 0)
    AND (FLargeFifo.IndexIn = 1) AND (FLargeFifo.IndexOut = 1)
    AND (FLargeStatus.SequenceId = 0) AND (FLargeStatus.DeletedSequenceId = 0)
    AND (FLargeStatus.LostEventCount = 0);
FOR Index := 1 TO LargeBufferLength DO
    FIsolationMatches := FIsolationMatches AND (FLargeEvents[Index].SequenceId = 0);
END_FOR;
END_METHOD

END_FUNCTION_BLOCK

// ---- SelfTests/TestCases/TestSuite_EventDelivery/Test_EventContent.TcPOU
{region 'Documentation'}
(*!
<summary>Verifies representative event payloads and producer-assigned identity through real publication.</summary>
<description>
Publishes a state transition, a failed Assertion and a Test Case aggregation. Expectations
state the required fields explicitly instead of constructing the expected event with the same FC.
Sequence and timestamp sentinels verify that the publisher assigns identity to its value copy.
Timestamp checks permit equal times; event ordering is determined only by SequenceId.
The real subject binds only local storage; expected findings remain in that storage.
Checking Assertions retain the outer selftest publisher. Each run reinitializes the subject.
</description>
*)
{endregion}
FUNCTION_BLOCK Test_EventContent EXTENDS TestCaseBase
VAR
    FSubject : EventBuffer;
    FEvents : ARRAY[1..BufferLength] OF ST_Event;
    FFifo : ST_FifoStatus;
    FBufferStatus : ST_EventBufferStatus;
    FPerformed : BOOL;
    FChecked : BOOL;
    FTransition : AssertTrue;
    FTransitionMatches : BOOL;
    FFinding : AssertTrue;
    FFindingMatches : BOOL;
    FAggregation : AssertTrue;
    FAggregationMatches : BOOL;
    FIdentity : AssertTrue;
    FIdentityMatches : BOOL;
    FValueCopy : AssertTrue;
    FValueCopyMatches : BOOL;
    FProjection : AssertTrue;
    FProjectionMatches : BOOL;
END_VAR
VAR CONSTANT
    BufferLength : UINT := 8;
    InputSequenceSentinel : UDINT := 999;
    InputTimestampSentinel : LINT := -1;
    TimestampResolutionNanoseconds : LINT := 100;
END_VAR

SUPER^();

{region 'Documentation'}
(*!
<summary>Contributes each checking Assertion once.</summary>
*)
{endregion}
METHOD PROTECTED AggregateResults
VAR_INPUT
    Aggregator : I_ResultAggregator; //! Borrowed result sink owned by the outer Test Case; add this test's checking Assertions without resetting or retaining the sink.
END_VAR
Aggregator.AddProvider(Provider := FTransition);
Aggregator.AddProvider(Provider := FFinding);
Aggregator.AddProvider(Provider := FAggregation);
Aggregator.AddProvider(Provider := FIdentity);
Aggregator.AddProvider(Provider := FValueCopy);
Aggregator.AddProvider(Provider := FProjection);
END_METHOD

{region 'Documentation'}
(*!
<summary>Requires all checking Assertions to be initialized.</summary>
*)
{endregion}
METHOD PROTECTED CheckInitialization : BOOL //! TRUE when the inherited initialization check and this concrete fixture check both accept the setup.
CheckInitialization := FALSE;
IF NOT SUPER^.CheckInitialization() THEN
    RETURN;
END_IF;

CheckInitialization := FTransition.IsInitialized
    AND FFinding.IsInitialized
    AND FAggregation.IsInitialized
    AND FIdentity.IsInitialized
    AND FValueCopy.IsInitialized
    AND FProjection.IsInitialized;
END_METHOD

{region 'Documentation'}
(*!
<summary>Initializes the checking Assertions for one test state.</summary>
*)
{endregion}
METHOD PROTECTED Configure
FPreparationStateCount := 0;
FTestStateCount := 1;
FTransition.Initialize(Parent := THIS^,
    AssertionName := 'Transition');
FFinding.Initialize(Parent := THIS^,
    AssertionName := 'Finding');
FAggregation.Initialize(Parent := THIS^,
    AssertionName := 'Aggregation');
FIdentity.Initialize(Parent := THIS^,
    AssertionName := 'Identity');
FValueCopy.Initialize(Parent := THIS^,
    AssertionName := 'ValueCopy');
FProjection.Initialize(Parent := THIS^,
    AssertionName := 'Projection');
END_METHOD

{region 'Documentation'}
(*!
<summary>Publishes three representative constructors and checks payload, identity and value-copy semantics.</summary>
*)
{endregion}
METHOD PRIVATE ExerciseBuffer
VAR
    Event : ST_Event;
    CaseStatus : ST_TestCaseStatus;
    WriteResult : INT;
    Index : UINT;
END_VAR
IF NOT FSubject.Initialize(Buffer := FEvents,
    FifoControl := FFifo,
    Status := FBufferStatus) THEN
    Error(Message := 'Local Event Buffer initialization failed.');
    RETURN;
END_IF;

Event := CreateStateTransitionEvent(OwnerScope := E_OwnerScope.TestCase,
    Name := 'Local.Suite.Case',
    ResourceName := 'Valve',
    StateOld := E_State.Idle,
    StateNew := E_State.Starting);
Event.SequenceId := InputSequenceSentinel;
Event.Timestamp := InputTimestampSentinel;
WriteResult := FSubject.PublishEvent(Event := Event);
FTransitionMatches := (WriteResult = 1)
    AND (FEvents[1].OwnerScope = E_OwnerScope.TestCase)
    AND (FEvents[1].EventType = E_EventType.StateTransition)
    AND (FEvents[1].Severity = E_EventSeverity.Info)
    AND (FEvents[1].Name = 'Local.Suite.Case') AND (FEvents[1].ResourceName = 'Valve')
    AND (FEvents[1].State = E_State.Starting) AND (FEvents[1].Result = E_Result.NotEvaluated)
    AND (FEvents[1].Message = 'State transition 10 -> 11');
FValueCopyMatches := (Event.SequenceId = InputSequenceSentinel)
    AND (Event.Timestamp = InputTimestampSentinel);

Event := CreateAssertionFailedEvent(Name := 'Local.Suite.Case.Position',
    ResourceName := 'Valve',
    State := E_State.Running,
    Message := 'Expected open, observed closed.');
WriteResult := FSubject.PublishEvent(Event := Event);
FFindingMatches := (WriteResult = 2)
    AND (FEvents[2].OwnerScope = E_OwnerScope.Assertion)
    AND (FEvents[2].EventType = E_EventType.Result)
    AND (FEvents[2].Severity = E_EventSeverity.Info)
    AND (FEvents[2].Name = 'Local.Suite.Case.Position') AND (FEvents[2].ResourceName = 'Valve')
    AND (FEvents[2].State = E_State.Running) AND (FEvents[2].Result = E_Result.Failed)
    AND (FEvents[2].Message = 'Expected open, observed closed.');
FValueCopyMatches := FValueCopyMatches AND (Event.SequenceId = 0) AND (Event.Timestamp = 0);

CaseStatus.Execution.State := E_State.Completing;
CaseStatus.Execution.Result := E_Result.Error;
CaseStatus.AssertionCountTotal := 6;
CaseStatus.AssertionCountPassed := 3;
CaseStatus.AssertionCountFailed := 2;
CaseStatus.AssertionCountError := 1;
CaseStatus.Runtime := T#123ms;
Event := CreateTestCaseAggregationEvent(Name := 'Local.Suite.Case',
    ResourceName := 'Valve',
    Status := CaseStatus);
WriteResult := FSubject.PublishEvent(Event := Event);
FAggregationMatches := (WriteResult = 3)
    AND (FEvents[3].OwnerScope = E_OwnerScope.TestCase)
    AND (FEvents[3].EventType = E_EventType.Aggregation)
    AND (FEvents[3].Severity = E_EventSeverity.Error)
    AND (FEvents[3].Name = 'Local.Suite.Case') AND (FEvents[3].ResourceName = 'Valve')
    AND (FEvents[3].State = E_State.Completing) AND (FEvents[3].Result = E_Result.Error)
    AND (FEvents[3].Message = '{"total":6,"passed":3,"failed":2,"error":1,"runtime":123}');
FValueCopyMatches := FValueCopyMatches AND (Event.SequenceId = 0) AND (Event.Timestamp = 0);

FIdentityMatches := TRUE;
FOR Index := 1 TO 3 DO
    FIdentityMatches := FIdentityMatches AND (FEvents[Index].SequenceId = UINT_TO_UDINT(Index))
        AND (FEvents[Index].Timestamp > 0)
        AND ((FEvents[Index].Timestamp MOD TimestampResolutionNanoseconds) = 0);
END_FOR;
FProjectionMatches := NOT FFifo.ConfigError AND NOT FFifo.IndexError
    AND NOT FFifo.BufferEmpty AND NOT FFifo.BufferFull AND NOT FFifo.BufferAlmostFull
    AND (FFifo.BufferLength = BufferLength) AND (FFifo.ElementCount = 3)
    AND (FFifo.IndexOut = 1) AND (FFifo.IndexIn = 4)
    AND (FSubject.FreeEntryCount = 4)
    AND (FBufferStatus.SequenceId = 3) AND (FBufferStatus.DeletedSequenceId = 0)
    AND (FBufferStatus.LostEventCount = 0);
END_METHOD

{region 'Documentation'}
(*!
<summary>Completes abort without asynchronous work.</summary>
*)
{endregion}
METHOD PROTECTED ProcessAbort
VAR_INPUT
    Enable : BOOL; //! Phase permission supplied by the owning Test Case; FALSE does not authorize progression, while observation may continue.
END_VAR
IF Enable THEN
    CompleteAbort();
END_IF;
END_METHOD

{region 'Documentation'}
(*!
<summary>Evaluates captured observations after the scenario has finished.</summary>
*)
{endregion}
METHOD PROTECTED ProcessAssertions
VAR_INPUT
    Enable : BOOL; //! Phase permission supplied by the owning Test Case; FALSE does not authorize progression, while observation may continue.
END_VAR
VAR
    Evaluate : BOOL;
END_VAR
Evaluate := Enable AND FPerformed;
FTransition(Enable := Evaluate,
    State := State,
    IN := FTransitionMatches);
FFinding(Enable := Evaluate,
    State := State,
    IN := FFindingMatches);
FAggregation(Enable := Evaluate,
    State := State,
    IN := FAggregationMatches);
FIdentity(Enable := Evaluate,
    State := State,
    IN := FIdentityMatches);
FValueCopy(Enable := Evaluate,
    State := State,
    IN := FValueCopyMatches);
FProjection(Enable := Evaluate,
    State := State,
    IN := FProjectionMatches);
IF Evaluate THEN
    FChecked := TRUE;
END_IF;
END_METHOD

{region 'Documentation'}
(*!
<summary>No Preparation phase is needed.</summary>
*)
{endregion}
METHOD PROTECTED ProcessPreparations
VAR_INPUT
    // SA0033: Required override without Preparation work.
    {attribute 'analysis' := '-33'}
    Enable : BOOL; //! Phase permission supplied by the owning Test Case; FALSE does not authorize progression, while observation may continue.
END_VAR
END_METHOD

{region 'Documentation'}
(*!
<summary>Resets observations and schedules a fresh subject initialization.</summary>
*)
{endregion}
METHOD PROTECTED ProcessReset
FPerformed := FALSE;
FChecked := FALSE;
FTransition.Reset();
FTransitionMatches := FALSE;
FFinding.Reset();
FFindingMatches := FALSE;
FAggregation.Reset();
FAggregationMatches := FALSE;
FIdentity.Reset();
FIdentityMatches := FALSE;
FValueCopy.Reset();
FValueCopyMatches := FALSE;
FProjection.Reset();
FProjectionMatches := FALSE;
CompleteReset();
END_METHOD

{region 'Documentation'}
(*!
<summary>Runs the bounded scenario once before Assertion evaluation.</summary>
*)
{endregion}
METHOD PROTECTED ProcessTests
VAR_INPUT
    Enable : BOOL; //! Phase permission supplied by the owning Test Case; FALSE does not authorize progression, while observation may continue.
END_VAR
IF NOT Enable THEN
    RETURN;
END_IF;
IF FChecked THEN
    CompleteTests();
    RETURN;
END_IF;

IF NOT FPerformed THEN
    ExerciseBuffer();
    FPerformed := TRUE;
END_IF;
END_METHOD

END_FUNCTION_BLOCK

// ---- SelfTests/TestCases/TestSuite_EventDelivery/Test_EventBufferFull.TcPOU
{region 'Documentation'}
(*!
<summary>Verifies full-buffer preservation, capacity diagnostics and loss accounting.</summary>
<description>
Four primary events fill four of five usable positions. The existing capacity diagnostic
occupies the fifth position. Two further publications must fail without overwriting any
stored event, while the assigned sequence and lost-event count advance.
The real subject binds only local storage; expected findings remain in that storage.
Checking Assertions retain the outer selftest publisher. Each run reinitializes the subject.
</description>
*)
{endregion}
FUNCTION_BLOCK Test_EventBufferFull EXTENDS TestCaseBase
VAR
    FSubject : EventBuffer;
    FEvents : ARRAY[1..BufferLength] OF ST_Event;
    FFifo : ST_FifoStatus;
    FBufferStatus : ST_EventBufferStatus;
    FPerformed : BOOL;
    FChecked : BOOL;
    FStoredEvents : ARRAY[1..BufferLength] OF ST_Event;
    FBeforeFull : AssertTrue;
    FBeforeFullMatches : BOOL;
    FFullProjection : AssertTrue;
    FFullProjectionMatches : BOOL;
    FCapacityDiagnostic : AssertTrue;
    FCapacityDiagnosticMatches : BOOL;
    FRejected : AssertTrue;
    FRejectedMatches : BOOL;
    FUnreadPreserved : AssertTrue;
    FUnreadPreservedMatches : BOOL;
    FLoss : AssertTrue;
    FLossMatches : BOOL;
END_VAR
VAR CONSTANT
    BufferLength : UINT := 6;
    PrimaryEventCount : UINT := 4;
END_VAR

SUPER^();

{region 'Documentation'}
(*!
<summary>Contributes each checking Assertion once.</summary>
*)
{endregion}
METHOD PROTECTED AggregateResults
VAR_INPUT
    Aggregator : I_ResultAggregator; //! Borrowed result sink owned by the outer Test Case; add this test's checking Assertions without resetting or retaining the sink.
END_VAR
Aggregator.AddProvider(Provider := FBeforeFull);
Aggregator.AddProvider(Provider := FFullProjection);
Aggregator.AddProvider(Provider := FCapacityDiagnostic);
Aggregator.AddProvider(Provider := FRejected);
Aggregator.AddProvider(Provider := FUnreadPreserved);
Aggregator.AddProvider(Provider := FLoss);
END_METHOD

{region 'Documentation'}
(*!
<summary>Requires all checking Assertions to be initialized.</summary>
*)
{endregion}
METHOD PROTECTED CheckInitialization : BOOL //! TRUE when the inherited initialization check and this concrete fixture check both accept the setup.
CheckInitialization := FALSE;
IF NOT SUPER^.CheckInitialization() THEN
    RETURN;
END_IF;

CheckInitialization := FBeforeFull.IsInitialized
    AND FFullProjection.IsInitialized
    AND FCapacityDiagnostic.IsInitialized
    AND FRejected.IsInitialized
    AND FUnreadPreserved.IsInitialized
    AND FLoss.IsInitialized;
END_METHOD

{region 'Documentation'}
(*!
<summary>Initializes the checking Assertions for one test state.</summary>
*)
{endregion}
METHOD PROTECTED Configure
FPreparationStateCount := 0;
FTestStateCount := 1;
FBeforeFull.Initialize(Parent := THIS^,
    AssertionName := 'BeforeFull');
FFullProjection.Initialize(Parent := THIS^,
    AssertionName := 'FullProjection');
FCapacityDiagnostic.Initialize(Parent := THIS^,
    AssertionName := 'CapacityDiagnostic');
FRejected.Initialize(Parent := THIS^,
    AssertionName := 'Rejected');
FUnreadPreserved.Initialize(Parent := THIS^,
    AssertionName := 'UnreadPreserved');
FLoss.Initialize(Parent := THIS^,
    AssertionName := 'Loss');
END_METHOD

{region 'Documentation'}
(*!
<summary>Fills the local buffer, captures its contents and attempts two rejected publications.</summary>
*)
{endregion}
METHOD PRIVATE ExerciseBuffer
VAR
    Event : ST_Event;
    WriteResult : INT;
    Index : UINT;
END_VAR
IF NOT FSubject.Initialize(Buffer := FEvents,
    FifoControl := FFifo,
    Status := FBufferStatus) THEN
    Error(Message := 'Local Event Buffer initialization failed.');
    RETURN;
END_IF;

FBeforeFullMatches := FFifo.BufferEmpty AND (FFifo.ElementCount = 0)
    AND (FSubject.FreeEntryCount = BufferLength - 1);
FOR Index := 1 TO PrimaryEventCount DO
    Event := CreateFrameworkEvent(Name := 'LocalFull',
        State := E_State.Running,
        Severity := E_EventSeverity.Info,
        Message := UINT_TO_STRING(Index));
    WriteResult := FSubject.PublishEvent(Event := Event);
    FBeforeFullMatches := FBeforeFullMatches AND (WriteResult = UINT_TO_INT(Index));
    IF Index < PrimaryEventCount THEN
        FBeforeFullMatches := FBeforeFullMatches AND NOT FFifo.BufferFull
            AND NOT FFifo.BufferAlmostFull AND (FFifo.ElementCount = Index)
            AND (FBufferStatus.SequenceId = UINT_TO_UDINT(Index))
            AND (FBufferStatus.LostEventCount = 0);
    END_IF;
END_FOR;

FFullProjectionMatches := FFifo.BufferFull AND NOT FFifo.BufferEmpty
    AND NOT FFifo.ConfigError AND NOT FFifo.IndexError
    AND (FFifo.BufferLength = BufferLength) AND (FFifo.ElementCount = BufferLength - 1)
    AND (FFifo.IndexOut = 1) AND (FFifo.IndexIn = BufferLength)
    AND (FSubject.FreeEntryCount = 0)
    AND (FBufferStatus.SequenceId = UINT_TO_UDINT(BufferLength - 1))
    AND (FBufferStatus.LostEventCount = 0);
FCapacityDiagnosticMatches := (FEvents[5].SequenceId = 5)
    AND (FEvents[5].OwnerScope = E_OwnerScope.Framework)
    AND (FEvents[5].EventType = E_EventType.Framework)
    AND (FEvents[5].Severity = E_EventSeverity.Error)
    AND (FEvents[5].Name = 'EventBuffer') AND (FEvents[5].Timestamp > 0);
FUnreadPreservedMatches := (FEvents[BufferLength].SequenceId = 0);
FOR Index := 1 TO PrimaryEventCount DO
    FUnreadPreservedMatches := FUnreadPreservedMatches
        AND (FEvents[Index].SequenceId = UINT_TO_UDINT(Index))
        AND (FEvents[Index].Name = 'LocalFull')
        AND (FEvents[Index].Message = UINT_TO_STRING(Index));
END_FOR;
FStoredEvents := FEvents;

Event := CreateFrameworkEvent(Name := 'Rejected',
    State := E_State.Running,
    Severity := E_EventSeverity.Info,
    Message := 'Must not replace an unread event.');
WriteResult := FSubject.PublishEvent(Event := Event);
FRejectedMatches := WriteResult = TO_INT(E_FifoResult.NoTransfer);
FLossMatches := (FBufferStatus.SequenceId = 6) AND (FBufferStatus.LostEventCount = 1);
WriteResult := FSubject.PublishEvent(Event := Event);
FRejectedMatches := FRejectedMatches AND (WriteResult = TO_INT(E_FifoResult.NoTransfer));
FLossMatches := FLossMatches AND (FBufferStatus.SequenceId = 7)
    AND (FBufferStatus.DeletedSequenceId = 0) AND (FBufferStatus.LostEventCount = 2)
    AND (FSubject.LostEventCount = 2);
FFullProjectionMatches := FFullProjectionMatches AND FFifo.BufferFull
    AND (FFifo.ElementCount = BufferLength - 1)
    AND (FFifo.IndexOut = 1) AND (FFifo.IndexIn = BufferLength)
    AND (FSubject.FreeEntryCount = 0);
FOR Index := 1 TO BufferLength DO
    FUnreadPreservedMatches := FUnreadPreservedMatches
        AND (FEvents[Index].SequenceId = FStoredEvents[Index].SequenceId)
        AND (FEvents[Index].Timestamp = FStoredEvents[Index].Timestamp)
        AND (FEvents[Index].OwnerScope = FStoredEvents[Index].OwnerScope)
        AND (FEvents[Index].EventType = FStoredEvents[Index].EventType)
        AND (FEvents[Index].Severity = FStoredEvents[Index].Severity)
        AND (FEvents[Index].Name = FStoredEvents[Index].Name)
        AND (FEvents[Index].ResourceName = FStoredEvents[Index].ResourceName)
        AND (FEvents[Index].State = FStoredEvents[Index].State)
        AND (FEvents[Index].Result = FStoredEvents[Index].Result)
        AND (FEvents[Index].Message = FStoredEvents[Index].Message);
END_FOR;
END_METHOD

{region 'Documentation'}
(*!
<summary>Completes abort without asynchronous work.</summary>
*)
{endregion}
METHOD PROTECTED ProcessAbort
VAR_INPUT
    Enable : BOOL; //! Phase permission supplied by the owning Test Case; FALSE does not authorize progression, while observation may continue.
END_VAR
IF Enable THEN
    CompleteAbort();
END_IF;
END_METHOD

{region 'Documentation'}
(*!
<summary>Evaluates captured observations after the scenario has finished.</summary>
*)
{endregion}
METHOD PROTECTED ProcessAssertions
VAR_INPUT
    Enable : BOOL; //! Phase permission supplied by the owning Test Case; FALSE does not authorize progression, while observation may continue.
END_VAR
VAR
    Evaluate : BOOL;
END_VAR
Evaluate := Enable AND FPerformed;
FBeforeFull(Enable := Evaluate,
    State := State,
    IN := FBeforeFullMatches);
FFullProjection(Enable := Evaluate,
    State := State,
    IN := FFullProjectionMatches);
FCapacityDiagnostic(Enable := Evaluate,
    State := State,
    IN := FCapacityDiagnosticMatches);
FRejected(Enable := Evaluate,
    State := State,
    IN := FRejectedMatches);
FUnreadPreserved(Enable := Evaluate,
    State := State,
    IN := FUnreadPreservedMatches);
FLoss(Enable := Evaluate,
    State := State,
    IN := FLossMatches);
IF Evaluate THEN
    FChecked := TRUE;
END_IF;
END_METHOD

{region 'Documentation'}
(*!
<summary>No Preparation phase is needed.</summary>
*)
{endregion}
METHOD PROTECTED ProcessPreparations
VAR_INPUT
    // SA0033: Required override without Preparation work.
    {attribute 'analysis' := '-33'}
    Enable : BOOL; //! Phase permission supplied by the owning Test Case; FALSE does not authorize progression, while observation may continue.
END_VAR
END_METHOD

{region 'Documentation'}
(*!
<summary>Resets observations and schedules a fresh subject initialization.</summary>
*)
{endregion}
METHOD PROTECTED ProcessReset
FPerformed := FALSE;
FChecked := FALSE;
FBeforeFull.Reset();
FBeforeFullMatches := FALSE;
FFullProjection.Reset();
FFullProjectionMatches := FALSE;
FCapacityDiagnostic.Reset();
FCapacityDiagnosticMatches := FALSE;
FRejected.Reset();
FRejectedMatches := FALSE;
FUnreadPreserved.Reset();
FUnreadPreservedMatches := FALSE;
FLoss.Reset();
FLossMatches := FALSE;
CompleteReset();
END_METHOD

{region 'Documentation'}
(*!
<summary>Runs the bounded scenario once before Assertion evaluation.</summary>
*)
{endregion}
METHOD PROTECTED ProcessTests
VAR_INPUT
    Enable : BOOL; //! Phase permission supplied by the owning Test Case; FALSE does not authorize progression, while observation may continue.
END_VAR
IF NOT Enable THEN
    RETURN;
END_IF;
IF FChecked THEN
    CompleteTests();
    RETURN;
END_IF;

IF NOT FPerformed THEN
    ExerciseBuffer();
    FPerformed := TRUE;
END_IF;
END_METHOD

END_FUNCTION_BLOCK

// ---- SelfTests/TestCases/TestSuite_EventDelivery/Test_EventRingOrder.TcPOU
{region 'Documentation'}
(*!
<summary>Verifies readable sequence order across the physical ring boundary and after draining.</summary>
<description>
Five events are published, then a valid watermark releases the first four. Four new events
occupy physical positions 6, 7, 8 and 1. Reading from IndexOut to IndexIn must yield
sequences 5 through 9, not physical array order. Valid deletion only arranges these states;
invalid watermark behavior belongs to separate tests. Draining does not reset the epoch.
The real subject binds only local storage; expected findings remain in that storage.
Checking Assertions retain the outer selftest publisher. Each run reinitializes the subject.
</description>
*)
{endregion}
FUNCTION_BLOCK Test_EventRingOrder EXTENDS TestCaseBase
VAR
    FSubject : EventBuffer;
    FEvents : ARRAY[1..BufferLength] OF ST_Event;
    FFifo : ST_FifoStatus;
    FBufferStatus : ST_EventBufferStatus;
    FPerformed : BOOL;
    FChecked : BOOL;
    FSetup : AssertTrue;
    FSetupMatches : BOOL;
    FWrappedProjection : AssertTrue;
    FWrappedProjectionMatches : BOOL;
    FReadableOrder : AssertTrue;
    FReadableOrderMatches : BOOL;
    FDrained : AssertTrue;
    FDrainedMatches : BOOL;
    FContinuedSequence : AssertTrue;
    FContinuedSequenceMatches : BOOL;
END_VAR
VAR CONSTANT
    BufferLength : UINT := 8;
    InitialEventCount : UINT := 5;
    LastWrappedSequence : UDINT := 9;
END_VAR

SUPER^();

{region 'Documentation'}
(*!
<summary>Contributes each checking Assertion once.</summary>
*)
{endregion}
METHOD PROTECTED AggregateResults
VAR_INPUT
    Aggregator : I_ResultAggregator; //! Borrowed result sink owned by the outer Test Case; add this test's checking Assertions without resetting or retaining the sink.
END_VAR
Aggregator.AddProvider(Provider := FSetup);
Aggregator.AddProvider(Provider := FWrappedProjection);
Aggregator.AddProvider(Provider := FReadableOrder);
Aggregator.AddProvider(Provider := FDrained);
Aggregator.AddProvider(Provider := FContinuedSequence);
END_METHOD

{region 'Documentation'}
(*!
<summary>Requires all checking Assertions to be initialized.</summary>
*)
{endregion}
METHOD PROTECTED CheckInitialization : BOOL //! TRUE when the inherited initialization check and this concrete fixture check both accept the setup.
CheckInitialization := FALSE;
IF NOT SUPER^.CheckInitialization() THEN
    RETURN;
END_IF;

CheckInitialization := FSetup.IsInitialized
    AND FWrappedProjection.IsInitialized
    AND FReadableOrder.IsInitialized
    AND FDrained.IsInitialized
    AND FContinuedSequence.IsInitialized;
END_METHOD

{region 'Documentation'}
(*!
<summary>Initializes the checking Assertions for one test state.</summary>
*)
{endregion}
METHOD PROTECTED Configure
FPreparationStateCount := 0;
FTestStateCount := 1;
FSetup.Initialize(Parent := THIS^,
    AssertionName := 'Setup');
FWrappedProjection.Initialize(Parent := THIS^,
    AssertionName := 'WrappedProjection');
FReadableOrder.Initialize(Parent := THIS^,
    AssertionName := 'ReadableOrder');
FDrained.Initialize(Parent := THIS^,
    AssertionName := 'Drained');
FContinuedSequence.Initialize(Parent := THIS^,
    AssertionName := 'ContinuedSequence');
END_METHOD

{region 'Documentation'}
(*!
<summary>Creates a wrapped readable range, drains it and publishes into the same epoch again.</summary>
*)
{endregion}
METHOD PRIVATE ExerciseBuffer
VAR
    Event : ST_Event;
    WriteResult : INT;
    Sequence : UDINT;
    DeleteSequence : UDINT;
    Index : UINT;
    Offset : UINT;
END_VAR
IF NOT FSubject.Initialize(Buffer := FEvents,
    FifoControl := FFifo,
    Status := FBufferStatus) THEN
    Error(Message := 'Local Event Buffer initialization failed.');
    RETURN;
END_IF;

FSetupMatches := TRUE;
FOR Sequence := 1 TO InitialEventCount DO
    Event := CreateFrameworkEvent(Name := 'LocalRing',
        State := E_State.Running,
        Severity := E_EventSeverity.Info,
        Message := UDINT_TO_STRING(Sequence));
    WriteResult := FSubject.PublishEvent(Event := Event);
    FSetupMatches := FSetupMatches AND (WriteResult = UDINT_TO_INT(Sequence));
END_FOR;
DeleteSequence := 4;
FSubject.ProcessDeleteRequest(SequenceId := DeleteSequence);
FSetupMatches := FSetupMatches AND (DeleteSequence = 0)
    AND (FFifo.IndexOut = 5) AND (FFifo.IndexIn = 6) AND (FFifo.ElementCount = 1)
    AND (FBufferStatus.SequenceId = 5) AND (FBufferStatus.DeletedSequenceId = 4)
    AND (FBufferStatus.LostEventCount = 0);

FOR Sequence := 6 TO LastWrappedSequence DO
    Event := CreateFrameworkEvent(Name := 'LocalRing',
        State := E_State.Running,
        Severity := E_EventSeverity.Info,
        Message := UDINT_TO_STRING(Sequence));
    WriteResult := FSubject.PublishEvent(Event := Event);
    FSetupMatches := FSetupMatches AND (WriteResult > TO_INT(E_FifoResult.NoTransfer));
END_FOR;
FWrappedProjectionMatches := NOT FFifo.ConfigError AND NOT FFifo.IndexError
    AND NOT FFifo.BufferEmpty AND NOT FFifo.BufferFull AND NOT FFifo.BufferAlmostFull
    AND (FFifo.BufferLength = BufferLength) AND (FFifo.ElementCount = 5)
    AND (FFifo.IndexOut = 5) AND (FFifo.IndexIn = 2)
    AND (FSubject.FreeEntryCount = 2)
    AND (FBufferStatus.SequenceId = LastWrappedSequence)
    AND (FBufferStatus.DeletedSequenceId = 4) AND (FBufferStatus.LostEventCount = 0);
FReadableOrderMatches := FALSE;
IF FWrappedProjectionMatches THEN
    // Table F traversal: start at IndexOut, wrap at BufferLength, exclude IndexIn.
    FReadableOrderMatches := TRUE;
    FOR Offset := 0 TO 4 DO
        Index := ((FFifo.IndexOut - 1 + Offset) MOD FFifo.BufferLength) + 1;
        FReadableOrderMatches := FReadableOrderMatches
            AND (FEvents[Index].SequenceId = UINT_TO_UDINT(5 + Offset))
            AND (FEvents[Index].Name = 'LocalRing')
            AND (FEvents[Index].Message = UINT_TO_STRING(5 + Offset));
    END_FOR;
END_IF;

DeleteSequence := LastWrappedSequence;
FSubject.ProcessDeleteRequest(SequenceId := DeleteSequence);
FDrainedMatches := (DeleteSequence = 0) AND FFifo.BufferEmpty AND NOT FFifo.BufferFull
    AND (FFifo.ElementCount = 0) AND (FFifo.IndexOut = 2) AND (FFifo.IndexIn = 2)
    AND (FSubject.FreeEntryCount = BufferLength - 1)
    AND (FBufferStatus.SequenceId = LastWrappedSequence)
    AND (FBufferStatus.DeletedSequenceId = LastWrappedSequence)
    AND (FBufferStatus.LostEventCount = 0);
FOR Index := 1 TO BufferLength DO
    FDrainedMatches := FDrainedMatches AND (FEvents[Index].SequenceId = 0);
END_FOR;

WriteResult := FSubject.PublishEvent(Event := CreateFrameworkEvent(Name := 'LocalRing',
    State := E_State.Running,
    Severity := E_EventSeverity.Info,
    Message := 'After drain'));
FContinuedSequenceMatches := (WriteResult = 2)
    AND (FEvents[2].SequenceId = LastWrappedSequence + 1)
    AND (FEvents[2].Message = 'After drain')
    AND NOT FFifo.BufferEmpty AND (FFifo.ElementCount = 1)
    AND (FFifo.IndexOut = 2) AND (FFifo.IndexIn = 3)
    AND (FBufferStatus.SequenceId = LastWrappedSequence + 1)
    AND (FBufferStatus.DeletedSequenceId = LastWrappedSequence)
    AND (FBufferStatus.LostEventCount = 0);
END_METHOD

{region 'Documentation'}
(*!
<summary>Completes abort without asynchronous work.</summary>
*)
{endregion}
METHOD PROTECTED ProcessAbort
VAR_INPUT
    Enable : BOOL; //! Phase permission supplied by the owning Test Case; FALSE does not authorize progression, while observation may continue.
END_VAR
IF Enable THEN
    CompleteAbort();
END_IF;
END_METHOD

{region 'Documentation'}
(*!
<summary>Evaluates captured observations after the scenario has finished.</summary>
*)
{endregion}
METHOD PROTECTED ProcessAssertions
VAR_INPUT
    Enable : BOOL; //! Phase permission supplied by the owning Test Case; FALSE does not authorize progression, while observation may continue.
END_VAR
VAR
    Evaluate : BOOL;
END_VAR
Evaluate := Enable AND FPerformed;
FSetup(Enable := Evaluate,
    State := State,
    IN := FSetupMatches);
FWrappedProjection(Enable := Evaluate,
    State := State,
    IN := FWrappedProjectionMatches);
FReadableOrder(Enable := Evaluate,
    State := State,
    IN := FReadableOrderMatches);
FDrained(Enable := Evaluate,
    State := State,
    IN := FDrainedMatches);
FContinuedSequence(Enable := Evaluate,
    State := State,
    IN := FContinuedSequenceMatches);
IF Evaluate THEN
    FChecked := TRUE;
END_IF;
END_METHOD

{region 'Documentation'}
(*!
<summary>No Preparation phase is needed.</summary>
*)
{endregion}
METHOD PROTECTED ProcessPreparations
VAR_INPUT
    // SA0033: Required override without Preparation work.
    {attribute 'analysis' := '-33'}
    Enable : BOOL; //! Phase permission supplied by the owning Test Case; FALSE does not authorize progression, while observation may continue.
END_VAR
END_METHOD

{region 'Documentation'}
(*!
<summary>Resets observations and schedules a fresh subject initialization.</summary>
*)
{endregion}
METHOD PROTECTED ProcessReset
FPerformed := FALSE;
FChecked := FALSE;
FSetup.Reset();
FSetupMatches := FALSE;
FWrappedProjection.Reset();
FWrappedProjectionMatches := FALSE;
FReadableOrder.Reset();
FReadableOrderMatches := FALSE;
FDrained.Reset();
FDrainedMatches := FALSE;
FContinuedSequence.Reset();
FContinuedSequenceMatches := FALSE;
CompleteReset();
END_METHOD

{region 'Documentation'}
(*!
<summary>Runs the bounded scenario once before Assertion evaluation.</summary>
*)
{endregion}
METHOD PROTECTED ProcessTests
VAR_INPUT
    Enable : BOOL; //! Phase permission supplied by the owning Test Case; FALSE does not authorize progression, while observation may continue.
END_VAR
IF NOT Enable THEN
    RETURN;
END_IF;
IF FChecked THEN
    CompleteTests();
    RETURN;
END_IF;

IF NOT FPerformed THEN
    ExerciseBuffer();
    FPerformed := TRUE;
END_IF;
END_METHOD

END_FUNCTION_BLOCK

// ---- SelfTests/TestCases/TestSuite_EventDelivery/Test_EventDeleteWatermarks.TcPOU
{region 'Documentation'}
(*!
<summary>Verifies zero, stale, valid and future deletion watermarks on local event storage.</summary>
<description>
Three retained events establish a prefix deletion. Zero and stale requests must not
move that prefix; future requests may append a diagnostic but must not release it.
The final stage repeats the future request on empty storage to distinguish rejection
from deleting the diagnostic that the rejection itself produces.
The real subject binds only local storage; expected findings remain in that storage.
Checking Assertions retain the outer selftest publisher. Each run reinitializes the subject.
</description>
*)
{endregion}
FUNCTION_BLOCK Test_EventDeleteWatermarks EXTENDS TestCaseBase
VAR
    FSubject : EventBuffer;
    FEvents : ARRAY[1..BufferLength] OF ST_Event;
    FFifo : ST_FifoStatus;
    FBufferStatus : ST_EventBufferStatus;
    FPerformed : BOOL;
    FChecked : BOOL;
    FZero : AssertTrue;
    FZeroMatches : BOOL;
    FPrefix : AssertTrue;
    FPrefixMatches : BOOL;
    FStale : AssertTrue;
    FStaleMatches : BOOL;
    FFuture : AssertTrue;
    FFutureMatches : BOOL;
    FDrained : AssertTrue;
    FDrainedMatches : BOOL;
    FEmptyFuture : AssertTrue;
    FEmptyFutureMatches : BOOL;
END_VAR
VAR CONSTANT
    BufferLength : UINT := 10;
END_VAR

SUPER^();

{region 'Documentation'}
(*!
<summary>Contributes each checking Assertion once.</summary>
*)
{endregion}
METHOD PROTECTED AggregateResults
VAR_INPUT
    Aggregator : I_ResultAggregator; //! Borrowed result sink owned by the outer Test Case; add this test's checking Assertions without resetting or retaining the sink.
END_VAR
Aggregator.AddProvider(Provider := FZero);
Aggregator.AddProvider(Provider := FPrefix);
Aggregator.AddProvider(Provider := FStale);
Aggregator.AddProvider(Provider := FFuture);
Aggregator.AddProvider(Provider := FDrained);
Aggregator.AddProvider(Provider := FEmptyFuture);
END_METHOD

{region 'Documentation'}
(*!
<summary>Drains to the last retained sequence and checks stale and future requests on empty storage.</summary>
*)
{endregion}
METHOD PRIVATE CheckEmptyBoundary
VAR
    Request : UDINT;
    Index : UINT;
END_VAR
Request := 4;
FSubject.ProcessDeleteRequest(SequenceId := Request);
FDrainedMatches := (Request = 0) AND FFifo.BufferEmpty AND (FFifo.ElementCount = 0)
    AND (FFifo.IndexOut = 5) AND (FFifo.IndexIn = 5)
    AND (FBufferStatus.SequenceId = 4) AND (FBufferStatus.DeletedSequenceId = 4);
Request := 4;
FSubject.ProcessDeleteRequest(SequenceId := Request);
FDrainedMatches := FDrainedMatches AND (Request = 0)
    AND FFifo.BufferEmpty AND (FFifo.ElementCount = 0)
    AND (FFifo.IndexOut = 5) AND (FFifo.IndexIn = 5)
    AND (FBufferStatus.SequenceId = 4) AND (FBufferStatus.DeletedSequenceId = 4)
    AND (FBufferStatus.LostEventCount = 0);
FOR Index := 1 TO BufferLength DO
    FDrainedMatches := FDrainedMatches AND (FEvents[Index].SequenceId = 0);
END_FOR;

Request := 5;
FSubject.ProcessDeleteRequest(SequenceId := Request);
FEmptyFutureMatches := (Request = 0) AND (FBufferStatus.DeletedSequenceId = 4)
    AND (FBufferStatus.SequenceId = 5) AND (FBufferStatus.LostEventCount = 0)
    AND NOT FFifo.BufferEmpty AND (FFifo.ElementCount = 1)
    AND (FFifo.IndexOut = 5) AND (FFifo.IndexIn = 6)
    AND (FEvents[5].SequenceId = 5) AND (FEvents[5].OwnerScope = E_OwnerScope.Framework)
    AND (FEvents[5].EventType = E_EventType.Framework)
    AND (FEvents[5].Severity = E_EventSeverity.Warning) AND (FEvents[5].Name = 'EventBuffer');
END_METHOD

{region 'Documentation'}
(*!
<summary>Requires all checking Assertions to be initialized.</summary>
*)
{endregion}
METHOD PROTECTED CheckInitialization : BOOL //! TRUE when the inherited initialization check and this concrete fixture check both accept the setup.
CheckInitialization := FALSE;
IF NOT SUPER^.CheckInitialization() THEN
    RETURN;
END_IF;

CheckInitialization := FZero.IsInitialized
    AND FPrefix.IsInitialized
    AND FStale.IsInitialized
    AND FFuture.IsInitialized
    AND FDrained.IsInitialized
    AND FEmptyFuture.IsInitialized;
END_METHOD

{region 'Documentation'}
(*!
<summary>Checks stale requests leave the suffix intact and a future request only appends a warning.</summary>
*)
{endregion}
METHOD PRIVATE CheckStaleAndFuture
VAR
    Request : UDINT;
    StaleSequence : UDINT;
END_VAR
FStaleMatches := TRUE;
FOR StaleSequence := 1 TO 2 DO
    Request := StaleSequence;
    FSubject.ProcessDeleteRequest(SequenceId := Request);
    FStaleMatches := FStaleMatches AND (Request = 0)
        AND (FFifo.ElementCount = 1) AND (FFifo.IndexOut = 3) AND (FFifo.IndexIn = 4)
        AND (FBufferStatus.SequenceId = 3) AND (FBufferStatus.DeletedSequenceId = 2)
        AND (FBufferStatus.LostEventCount = 0)
        AND (FEvents[3].SequenceId = 3) AND (FEvents[3].Message = '3');
END_FOR;

Request := 100;
FSubject.ProcessDeleteRequest(SequenceId := Request);
FFutureMatches := (Request = 0) AND (FBufferStatus.DeletedSequenceId = 2)
    AND (FBufferStatus.SequenceId = 4) AND (FBufferStatus.LostEventCount = 0)
    AND (FFifo.ElementCount = 2) AND (FFifo.IndexOut = 3) AND (FFifo.IndexIn = 5)
    AND (FEvents[3].SequenceId = 3) AND (FEvents[3].Name = 'LocalDelete')
    AND (FEvents[3].Message = '3')
    AND (FEvents[4].SequenceId = 4) AND (FEvents[4].OwnerScope = E_OwnerScope.Framework)
    AND (FEvents[4].EventType = E_EventType.Framework)
    AND (FEvents[4].Severity = E_EventSeverity.Warning) AND (FEvents[4].Name = 'EventBuffer');
END_METHOD

{region 'Documentation'}
(*!
<summary>Checks zero requests on empty and occupied storage, followed by exact prefix deletion.</summary>
*)
{endregion}
METHOD PRIVATE CheckZeroAndPrefix
VAR
    Request : UDINT;
    Index : UINT;
    WriteResult : INT;
END_VAR
Request := 0;
FSubject.ProcessDeleteRequest(SequenceId := Request);
FZeroMatches := (Request = 0) AND FFifo.BufferEmpty AND (FFifo.ElementCount = 0)
    AND (FFifo.IndexIn = 1) AND (FFifo.IndexOut = 1)
    AND (FBufferStatus.SequenceId = 0) AND (FBufferStatus.DeletedSequenceId = 0)
    AND (FBufferStatus.LostEventCount = 0);
FOR Index := 1 TO 3 DO
    WriteResult := FSubject.PublishEvent(Event := CreateFrameworkEvent(Name := 'LocalDelete',
        State := E_State.Running,
        Severity := E_EventSeverity.Info,
        Message := UINT_TO_STRING(Index)));
    FZeroMatches := FZeroMatches AND (WriteResult = UINT_TO_INT(Index));
END_FOR;
Request := 0;
FSubject.ProcessDeleteRequest(SequenceId := Request);
FZeroMatches := FZeroMatches AND (Request = 0)
    AND (FFifo.ElementCount = 3) AND (FFifo.IndexOut = 1) AND (FFifo.IndexIn = 4)
    AND (FBufferStatus.SequenceId = 3) AND (FBufferStatus.DeletedSequenceId = 0)
    AND (FBufferStatus.LostEventCount = 0);
FOR Index := 1 TO 3 DO
    FZeroMatches := FZeroMatches AND (FEvents[Index].SequenceId = UINT_TO_UDINT(Index))
        AND (FEvents[Index].Name = 'LocalDelete') AND (FEvents[Index].Message = UINT_TO_STRING(Index));
END_FOR;

Request := 2;
FSubject.ProcessDeleteRequest(SequenceId := Request);
FPrefixMatches := (Request = 0) AND (FBufferStatus.DeletedSequenceId = 2)
    AND (FBufferStatus.SequenceId = 3) AND (FBufferStatus.LostEventCount = 0)
    AND (FFifo.ElementCount = 1) AND (FFifo.IndexOut = 3) AND (FFifo.IndexIn = 4)
    AND (FEvents[3].SequenceId = 3) AND (FEvents[3].Name = 'LocalDelete')
    AND (FEvents[3].Message = '3');
FOR Index := 1 TO 2 DO
    FPrefixMatches := FPrefixMatches AND (FEvents[Index].SequenceId = 0)
        AND (FEvents[Index].Timestamp = 0) AND (FEvents[Index].Name = '')
        AND (FEvents[Index].Message = '');
END_FOR;
END_METHOD

{region 'Documentation'}
(*!
<summary>Initializes the checking Assertions for one test state.</summary>
*)
{endregion}
METHOD PROTECTED Configure
FPreparationStateCount := 0;
FTestStateCount := 1;
FZero.Initialize(Parent := THIS^,
    AssertionName := 'Zero');
FPrefix.Initialize(Parent := THIS^,
    AssertionName := 'Prefix');
FStale.Initialize(Parent := THIS^,
    AssertionName := 'Stale');
FFuture.Initialize(Parent := THIS^,
    AssertionName := 'Future');
FDrained.Initialize(Parent := THIS^,
    AssertionName := 'Drained');
FEmptyFuture.Initialize(Parent := THIS^,
    AssertionName := 'EmptyFuture');
END_METHOD

{region 'Documentation'}
(*!
<summary>Initializes a local subject, then exercises the watermark boundaries in order.</summary>
*)
{endregion}
METHOD PRIVATE ExerciseBuffer
IF NOT FSubject.Initialize(Buffer := FEvents,
    FifoControl := FFifo,
    Status := FBufferStatus) THEN
    Error(Message := 'Local Event Buffer initialization failed.');
    RETURN;
END_IF;

CheckZeroAndPrefix();
CheckStaleAndFuture();
CheckEmptyBoundary();
END_METHOD

{region 'Documentation'}
(*!
<summary>Completes abort without asynchronous work.</summary>
*)
{endregion}
METHOD PROTECTED ProcessAbort
VAR_INPUT
    Enable : BOOL; //! Phase permission supplied by the owning Test Case; FALSE does not authorize progression, while observation may continue.
END_VAR
IF Enable THEN
    CompleteAbort();
END_IF;
END_METHOD

{region 'Documentation'}
(*!
<summary>Evaluates captured observations after the scenario has finished.</summary>
*)
{endregion}
METHOD PROTECTED ProcessAssertions
VAR_INPUT
    Enable : BOOL; //! Phase permission supplied by the owning Test Case; FALSE does not authorize progression, while observation may continue.
END_VAR
VAR
    Evaluate : BOOL;
END_VAR
Evaluate := Enable AND FPerformed;
FZero(Enable := Evaluate,
    State := State,
    IN := FZeroMatches);
FPrefix(Enable := Evaluate,
    State := State,
    IN := FPrefixMatches);
FStale(Enable := Evaluate,
    State := State,
    IN := FStaleMatches);
FFuture(Enable := Evaluate,
    State := State,
    IN := FFutureMatches);
FDrained(Enable := Evaluate,
    State := State,
    IN := FDrainedMatches);
FEmptyFuture(Enable := Evaluate,
    State := State,
    IN := FEmptyFutureMatches);
IF Evaluate THEN
    FChecked := TRUE;
END_IF;
END_METHOD

{region 'Documentation'}
(*!
<summary>No Preparation phase is needed.</summary>
*)
{endregion}
METHOD PROTECTED ProcessPreparations
VAR_INPUT
    // SA0033: Required override without Preparation work.
    {attribute 'analysis' := '-33'}
    Enable : BOOL; //! Phase permission supplied by the owning Test Case; FALSE does not authorize progression, while observation may continue.
END_VAR
END_METHOD

{region 'Documentation'}
(*!
<summary>Resets observations and schedules a fresh subject initialization.</summary>
*)
{endregion}
METHOD PROTECTED ProcessReset
FPerformed := FALSE;
FChecked := FALSE;
FZero.Reset();
FZeroMatches := FALSE;
FPrefix.Reset();
FPrefixMatches := FALSE;
FStale.Reset();
FStaleMatches := FALSE;
FFuture.Reset();
FFutureMatches := FALSE;
FDrained.Reset();
FDrainedMatches := FALSE;
FEmptyFuture.Reset();
FEmptyFutureMatches := FALSE;
CompleteReset();
END_METHOD

{region 'Documentation'}
(*!
<summary>Runs the bounded scenario once before Assertion evaluation.</summary>
*)
{endregion}
METHOD PROTECTED ProcessTests
VAR_INPUT
    Enable : BOOL; //! Phase permission supplied by the owning Test Case; FALSE does not authorize progression, while observation may continue.
END_VAR
IF NOT Enable THEN
    RETURN;
END_IF;
IF FChecked THEN
    CompleteTests();
    RETURN;
END_IF;

IF NOT FPerformed THEN
    ExerciseBuffer();
    FPerformed := TRUE;
END_IF;
END_METHOD

END_FUNCTION_BLOCK

// ---- SelfTests/TestCases/TestSuite_EventDelivery/Test_EventDeleteWrappedFull.TcPOU
{region 'Documentation'}
(*!
<summary>Verifies prefix deletion from full storage before and after a physical ring wrap.</summary>
<description>
Six primary events plus the capacity diagnostic fill seven usable slots. Deleting through
sequence 4 permits three further primary events and a new capacity diagnostic. The next
watermark is 9, beyond the physical upper index 8: it removes sequences 5 through 9
across the ring boundary while retaining sequences 10 and 11.
The real subject binds only local storage; expected findings remain in that storage.
Checking Assertions retain the outer selftest publisher. Each run reinitializes the subject.
</description>
*)
{endregion}
FUNCTION_BLOCK Test_EventDeleteWrappedFull EXTENDS TestCaseBase
VAR
    FSubject : EventBuffer;
    FEvents : ARRAY[1..BufferLength] OF ST_Event;
    FFifo : ST_FifoStatus;
    FBufferStatus : ST_EventBufferStatus;
    FPerformed : BOOL;
    FChecked : BOOL;
    FInitialFull : AssertTrue;
    FInitialFullMatches : BOOL;
    FFullPrefix : AssertTrue;
    FFullPrefixMatches : BOOL;
    FWrappedFull : AssertTrue;
    FWrappedFullMatches : BOOL;
    FWrappedPrefix : AssertTrue;
    FWrappedPrefixMatches : BOOL;
    FDrained : AssertTrue;
    FDrainedMatches : BOOL;
END_VAR
VAR CONSTANT
    BufferLength : UINT := 8;
END_VAR

SUPER^();

{region 'Documentation'}
(*!
<summary>Contributes each checking Assertion once.</summary>
*)
{endregion}
METHOD PROTECTED AggregateResults
VAR_INPUT
    Aggregator : I_ResultAggregator; //! Borrowed result sink owned by the outer Test Case; add this test's checking Assertions without resetting or retaining the sink.
END_VAR
Aggregator.AddProvider(Provider := FInitialFull);
Aggregator.AddProvider(Provider := FFullPrefix);
Aggregator.AddProvider(Provider := FWrappedFull);
Aggregator.AddProvider(Provider := FWrappedPrefix);
Aggregator.AddProvider(Provider := FDrained);
END_METHOD

{region 'Documentation'}
(*!
<summary>Requires all checking Assertions to be initialized.</summary>
*)
{endregion}
METHOD PROTECTED CheckInitialization : BOOL //! TRUE when the inherited initialization check and this concrete fixture check both accept the setup.
CheckInitialization := FALSE;
IF NOT SUPER^.CheckInitialization() THEN
    RETURN;
END_IF;

CheckInitialization := FInitialFull.IsInitialized
    AND FFullPrefix.IsInitialized
    AND FWrappedFull.IsInitialized
    AND FWrappedPrefix.IsInitialized
    AND FDrained.IsInitialized;
END_METHOD

{region 'Documentation'}
(*!
<summary>Initializes the checking Assertions for one test state.</summary>
*)
{endregion}
METHOD PROTECTED Configure
FPreparationStateCount := 0;
FTestStateCount := 1;
FInitialFull.Initialize(Parent := THIS^,
    AssertionName := 'InitialFull');
FFullPrefix.Initialize(Parent := THIS^,
    AssertionName := 'FullPrefix');
FWrappedFull.Initialize(Parent := THIS^,
    AssertionName := 'WrappedFull');
FWrappedPrefix.Initialize(Parent := THIS^,
    AssertionName := 'WrappedPrefix');
FDrained.Initialize(Parent := THIS^,
    AssertionName := 'Drained');
END_METHOD

{region 'Documentation'}
(*!
<summary>Uses sequence 9 rather than a physical index, preserves the suffix and then drains it.</summary>
*)
{endregion}
METHOD PRIVATE DeleteWrappedPrefix
VAR
    Request : UDINT;
    Index : UINT;
END_VAR
Request := 9;
FSubject.ProcessDeleteRequest(SequenceId := Request);
FWrappedPrefixMatches := (Request = 0) AND NOT FFifo.BufferFull AND NOT FFifo.BufferEmpty
    AND (FFifo.ElementCount = 2) AND (FFifo.IndexOut = 2) AND (FFifo.IndexIn = 4)
    AND (FBufferStatus.DeletedSequenceId = 9) AND (FBufferStatus.SequenceId = 11)
    AND (FBufferStatus.LostEventCount = 0)
    AND (FEvents[1].SequenceId = 0) AND (FEvents[1].Timestamp = 0)
    AND (FEvents[1].Name = '') AND (FEvents[1].Message = '')
    AND (FEvents[2].SequenceId = 10) AND (FEvents[2].Name = 'LocalWrappedDelete')
    AND (FEvents[2].Message = '10')
    AND (FEvents[3].SequenceId = 11) AND (FEvents[3].Name = 'EventBuffer');
FOR Index := 5 TO 8 DO
    FWrappedPrefixMatches := FWrappedPrefixMatches AND (FEvents[Index].SequenceId = 0)
        AND (FEvents[Index].Timestamp = 0) AND (FEvents[Index].Name = '') AND (FEvents[Index].Message = '');
END_FOR;

Request := 11;
FSubject.ProcessDeleteRequest(SequenceId := Request);
FDrainedMatches := (Request = 0) AND FFifo.BufferEmpty AND NOT FFifo.BufferFull
    AND (FFifo.ElementCount = 0) AND (FFifo.IndexOut = 4) AND (FFifo.IndexIn = 4)
    AND (FSubject.FreeEntryCount = 7)
    AND (FBufferStatus.SequenceId = 11) AND (FBufferStatus.DeletedSequenceId = 11)
    AND (FBufferStatus.LostEventCount = 0);
FOR Index := 1 TO BufferLength DO
    FDrainedMatches := FDrainedMatches AND (FEvents[Index].SequenceId = 0);
END_FOR;
END_METHOD

{region 'Documentation'}
(*!
<summary>Creates a full ring, advances its head, fills across wrap and deletes the selected prefix.</summary>
*)
{endregion}
METHOD PRIVATE ExerciseBuffer
IF NOT FSubject.Initialize(Buffer := FEvents,
    FifoControl := FFifo,
    Status := FBufferStatus) THEN
    Error(Message := 'Local Event Buffer initialization failed.');
    RETURN;
END_IF;

FillAndDeletePrefix();
FillWrappedRange();
DeleteWrappedPrefix();
END_METHOD

{region 'Documentation'}
(*!
<summary>Fills seven usable positions and releases exactly the first four events.</summary>
*)
{endregion}
METHOD PRIVATE FillAndDeletePrefix
VAR
    Index : UINT;
    Request : UDINT;
    WriteResult : INT;
END_VAR
FInitialFullMatches := TRUE;
FOR Index := 1 TO 6 DO
    WriteResult := FSubject.PublishEvent(Event := CreateFrameworkEvent(Name := 'LocalWrappedDelete',
        State := E_State.Running,
        Severity := E_EventSeverity.Info,
        Message := UINT_TO_STRING(Index)));
    FInitialFullMatches := FInitialFullMatches AND (WriteResult = UINT_TO_INT(Index));
END_FOR;
FInitialFullMatches := FInitialFullMatches AND FFifo.BufferFull
    AND (FFifo.ElementCount = 7) AND (FFifo.IndexOut = 1) AND (FFifo.IndexIn = 8)
    AND (FBufferStatus.SequenceId = 7) AND (FBufferStatus.DeletedSequenceId = 0)
    AND (FBufferStatus.LostEventCount = 0) AND (FEvents[7].SequenceId = 7)
    AND (FEvents[7].Name = 'EventBuffer');

Request := 4;
FSubject.ProcessDeleteRequest(SequenceId := Request);
FFullPrefixMatches := (Request = 0) AND NOT FFifo.BufferFull
    AND (FFifo.ElementCount = 3) AND (FFifo.IndexOut = 5) AND (FFifo.IndexIn = 8)
    AND (FBufferStatus.DeletedSequenceId = 4) AND (FBufferStatus.SequenceId = 7)
    AND (FBufferStatus.LostEventCount = 0);
FOR Index := 1 TO 4 DO
    FFullPrefixMatches := FFullPrefixMatches AND (FEvents[Index].SequenceId = 0)
        AND (FEvents[Index].Timestamp = 0) AND (FEvents[Index].Name = '') AND (FEvents[Index].Message = '');
END_FOR;
FOR Index := 5 TO 7 DO
    FFullPrefixMatches := FFullPrefixMatches AND (FEvents[Index].SequenceId = UINT_TO_UDINT(Index));
END_FOR;
END_METHOD

{region 'Documentation'}
(*!
<summary>Fills positions 8, 1 and 2; the capacity diagnostic occupies position 3.</summary>
*)
{endregion}
METHOD PRIVATE FillWrappedRange
VAR
    Sequence : UDINT;
    WriteResult : INT;
END_VAR
FWrappedFullMatches := TRUE;
FOR Sequence := 8 TO 10 DO
    WriteResult := FSubject.PublishEvent(Event := CreateFrameworkEvent(Name := 'LocalWrappedDelete',
        State := E_State.Running,
        Severity := E_EventSeverity.Info,
        Message := UDINT_TO_STRING(Sequence)));
    FWrappedFullMatches := FWrappedFullMatches AND (WriteResult > TO_INT(E_FifoResult.NoTransfer));
END_FOR;
FWrappedFullMatches := FWrappedFullMatches AND FFifo.BufferFull
    AND (FFifo.ElementCount = 7) AND (FFifo.IndexOut = 5) AND (FFifo.IndexIn = 4)
    AND (FBufferStatus.SequenceId = 11) AND (FBufferStatus.DeletedSequenceId = 4)
    AND (FBufferStatus.LostEventCount = 0)
    AND (FEvents[8].SequenceId = 8) AND (FEvents[1].SequenceId = 9)
    AND (FEvents[2].SequenceId = 10) AND (FEvents[3].SequenceId = 11)
    AND (FEvents[3].Name = 'EventBuffer') AND (FEvents[3].Severity = E_EventSeverity.Error);
END_METHOD

{region 'Documentation'}
(*!
<summary>Completes abort without asynchronous work.</summary>
*)
{endregion}
METHOD PROTECTED ProcessAbort
VAR_INPUT
    Enable : BOOL; //! Phase permission supplied by the owning Test Case; FALSE does not authorize progression, while observation may continue.
END_VAR
IF Enable THEN
    CompleteAbort();
END_IF;
END_METHOD

{region 'Documentation'}
(*!
<summary>Evaluates captured observations after the scenario has finished.</summary>
*)
{endregion}
METHOD PROTECTED ProcessAssertions
VAR_INPUT
    Enable : BOOL; //! Phase permission supplied by the owning Test Case; FALSE does not authorize progression, while observation may continue.
END_VAR
VAR
    Evaluate : BOOL;
END_VAR
Evaluate := Enable AND FPerformed;
FInitialFull(Enable := Evaluate,
    State := State,
    IN := FInitialFullMatches);
FFullPrefix(Enable := Evaluate,
    State := State,
    IN := FFullPrefixMatches);
FWrappedFull(Enable := Evaluate,
    State := State,
    IN := FWrappedFullMatches);
FWrappedPrefix(Enable := Evaluate,
    State := State,
    IN := FWrappedPrefixMatches);
FDrained(Enable := Evaluate,
    State := State,
    IN := FDrainedMatches);
IF Evaluate THEN
    FChecked := TRUE;
END_IF;
END_METHOD

{region 'Documentation'}
(*!
<summary>No Preparation phase is needed.</summary>
*)
{endregion}
METHOD PROTECTED ProcessPreparations
VAR_INPUT
    // SA0033: Required override without Preparation work.
    {attribute 'analysis' := '-33'}
    Enable : BOOL; //! Phase permission supplied by the owning Test Case; FALSE does not authorize progression, while observation may continue.
END_VAR
END_METHOD

{region 'Documentation'}
(*!
<summary>Resets observations and schedules a fresh subject initialization.</summary>
*)
{endregion}
METHOD PROTECTED ProcessReset
FPerformed := FALSE;
FChecked := FALSE;
FInitialFull.Reset();
FInitialFullMatches := FALSE;
FFullPrefix.Reset();
FFullPrefixMatches := FALSE;
FWrappedFull.Reset();
FWrappedFullMatches := FALSE;
FWrappedPrefix.Reset();
FWrappedPrefixMatches := FALSE;
FDrained.Reset();
FDrainedMatches := FALSE;
CompleteReset();
END_METHOD

{region 'Documentation'}
(*!
<summary>Runs the bounded scenario once before Assertion evaluation.</summary>
*)
{endregion}
METHOD PROTECTED ProcessTests
VAR_INPUT
    Enable : BOOL; //! Phase permission supplied by the owning Test Case; FALSE does not authorize progression, while observation may continue.
END_VAR
IF NOT Enable THEN
    RETURN;
END_IF;
IF FChecked THEN
    CompleteTests();
    RETURN;
END_IF;

IF NOT FPerformed THEN
    ExerciseBuffer();
    FPerformed := TRUE;
END_IF;
END_METHOD

END_FUNCTION_BLOCK

